      def clipWhenLowerLimitIsLessThanHigher(outputScaledValue, outputRange):
          if (outputScaledValue < outputRange[0]):
              return outputRange[0]
          elif (outputScaledValue > outputRange[1]):
              return outputRange[1]
          else:
              return outputScaledValue
          end
      end

      slope = computeSlope(rawRange, scaledRange)
      intercept = computeIntercept(slope, rawRange, scaledRange)
      scaledValue = slope * value + intercept
      return clipScaledValue(scaledValue, scaledRange)
  end

  def limit(value, range):
      return scale(value, range, range)
  end


  rq_init_comm_if_connected(9, "1")
  rq_init_comm_if_connected(2, "2")
  rq_init_comm_if_connected(3, "3")
  rq_init_comm_if_connected(4, "4")
  rq_print_connected_grippers()
  rq_gripper_communication_thread = run rq_gripper_communication()
  set_closed_norm(97.6470588235294, 1)
  set_open_norm(1.1764705882352942, 1)
  set_closed_mm(0.0, 1)
  set_open_mm(53.0, 1)
  set_closed_norm(100.0, 2)
  set_open_norm(0.0, 2)
  set_closed_mm(0.0, 2)
  set_open_mm(50.0, 2)
  set_closed_norm(100.0, 3)
  set_open_norm(0.0, 3)
  set_closed_mm(0.0, 3)
  set_open_mm(50.0, 3)
  set_closed_norm(100.0, 4)
  set_open_norm(0.0, 4)
  set_closed_mm(0.0, 4)
  set_open_mm(50.0, 4)
  rq_current_limit_enabled = False
  while(not rq_gripper_communication_thread_started):
      sync()
  end
  # end: URCap Installation Node
  # begin: URCap Installation Node
  #   Source: OPC UA, 2.0.2, Rocketfarm AS
  #   Type: OPC UA
  global opcua_daemon = rpc_factory("xmlrpc", "http://127.0.0.1:40409/RPC2")
  def opcua_client_connect(address):
  return opcua_daemon.client_connect(address)
  end
  def opcua_client_get_id(client_name):
  return opcua_daemon.client_get_id(client_name)
  end
  def opcua_client_try_connect(client_id):
  opcua_result = False
  if (opcua_daemon.client_connect(client_id)):
  sleep(0.01)
  opcua_result = opcua_daemon.client_is_connected(client_id)
  opcua_retry = 10
  while ( (not opcua_result) and (opcua_retry > 0) ):
  sleep(0.1)
  opcua_result = opcua_daemon.client_is_connected(client_id)
  opcua_retry = opcua_retry - 1
  end
  end
  return opcua_result
  end
  def opcua_client_disconnect(client_id):
  return opcua_daemon.client_disconnect(client_id)
  end
  def opcua_client_is_connected(client_id):
  return opcua_daemon.client_is_connected(client_id)
  end
  def opcua_client_read_byid(client_id, namespace_id, variable_id):
  return opcua_daemon.client_read_variable_by_id(client_id, namespace_id, variable_id)
  end
  def opcua_client_read_byname(client_id, namespace_id, variable_name):
  return opcua_daemon.client_read_variable_by_name(client_id, namespace_id, variable_name)
  end
  def opcua_client_write_byid(client_id, namespace_id, variable_id, variable_value):
  return opcua_daemon.client_write_variable_by_id(client_id, namespace_id, variable_id, variable_value)
  end
  def opcua_client_write_byname(client_id, namespace_id, variable_name, variable_value):
  return opcua_daemon.client_write_variable_by_name(client_id, namespace_id, variable_name, variable_value)
  end
  def opcua_client_last_error(client_id):
  return opcua_daemon.client_get_last_error(client_id)
  end
  def opcua_server_read_byname(variable_name):
  return opcua_daemon.server_read_variable_by_name(variable_name)
  end
  def opcua_server_write_byname(variable_name, variable_value):
  return opcua_daemon.server_write_variable_by_name(variable_name, variable_value)
  end
  def opcua_server_last_error():
  return opcua_daemon.server_get_last_error()
  end
  def opcua_error_to_string(errorCode):
  return opcua_daemon.error_code_to_string(errorCode)
  end
  # end: URCap Installation Node
  global AMR_Position=struct(position_identifier=0, x1=0, x2=0, y1=0, y2=0, theta1=0, theta2=0)
  global CAM_Pose=p[0,0,0,0,0,0]
  global CAM_Relation=""
  global CMD_Abort=  False
  global CMD_Clear=  False
  global CMD_Reset=  False
  global CMD_Start=  False
  global CMD_Suspend=  False
  global CMD_Unhold=  False
  global CMD_Unsuspend=  False
  global CNT_Rack_Output=0
  global FNC_Freedrive=  False
  global PRC_TubCounter=0
  global STP=0
  global easyPickCount=0
  global easyPickCount_4=0
  global easyPickCount_6=0
  global easyPickCount_7=0
  global easyPickNoObj=0
  global easyPickNoObj_4=0
  global easyPickNoObj_6=0
  global easyPickNoObj_7=0
  global easyPickParts=0
  global easyPickParts_4=0
  global easyPickParts_6=0
  global easyPickParts_7=0
  global Container_mid_1_p=p[-.379239199143, -.127191311915, .299999999998, .000000000046, -.000000000021, -1.247199999994]
  global Container_mid_1_q=[-2.477408934449926, -1.2969853503591224, -1.875639182904262, -1.539621866126728, 1.5731943360401213, -2.8009955944022717]
  global Container_capt_p=p[-.525590029047, .407247642794, .411588185841, -.000000000107, .000000000065, -2.896148821900]
  global Container_capt_q=[-3.5968351615224767, -2.0050156108707204, -0.8176271154495112, -1.8895759482008394, 1.5730967555598792, -2.2743681102957645]
  global Waypoint_51_p=p[-.335468094724, -.217855817953, .299999999998, .000000000047, -.000000000014, -.994837065669]
  global Waypoint_51_q=[-2.2250460001249586, -1.2969853503591224, -1.875639182904262, -1.539621866126728, 1.573194336040121, -2.800995594402271]
  global Waypoint_13_p=p[-.479450777041, .284140798427, .125270103493, -.276792173670, 2.098433187455, -2.121256516887]
  global Waypoint_13_q=[-2.8915050665484827, -1.9549266300597132, -2.2318272590637207, -1.6654960117735804, 0.020810842514038086, -0.4019392172442835]
  global Waypoint_70_p=p[-.472820924464, .292439826304, .207418370234, -.259787347864, -2.053484648504, 2.070709755662]
  global Waypoint_70_q=[-2.969927421603815, -2.07168115810532, -1.6835546062719366, -2.4953958198513964, 0.4489790927922641, -0.005578998612037367]
  global Waypoint_2_p=p[-.312961047461, -.152991312519, .223609826854, -.745314530454, -1.713873240489, 1.673341715282]
  global Waypoint_2_q=[-2.3560472170459192, -2.183784624139303, -1.4583134651184082, -2.6435262165465296, 1.6522362232208252, 0.043451953679323196]
  global Waypoint_3_p=p[-.113749865836, -.390110151572, .317307487562, -.519383711706, -.839884211339, 1.756868173041]
  global Waypoint_3_q=[-1.8909733931170862, -1.720626016656393, -1.5115610361099243, -2.1240560017027796, 2.1809096336364746, 0.7227501273155212]
  global Waypoint_15_p=p[.029144035010, -.436802470887, .327885032028, -.521560953301, -.623641814548, 1.862659450154]
  global Waypoint_15_q=[-1.564817253743307, -1.556895188321807, -1.6826975345611572, -1.6944714985289515, 2.2362685203552246, 1.117417335510254]
  global Waypoint_14_p=p[.068712235638, -.569419545175, .285215357659, -.679242949116, -.712065334485, 1.394044574094]
  global Waypoint_14_q=[-1.5731792953485346, -1.8029235103747094, -1.6781008808776736, -1.2218450646111982, 2.4719572998240125, 1.6394218026856375]
  global Waypoint_4_p=p[-.047220457210, -.557624911767, .136370962514, -.679242949107, -.712065334475, 1.394044574096]
  global Waypoint_4_q=[-1.7740079055958748, -2.0023561428872334, -1.7577251142892676, -1.18903287716154, 2.4487287370345143, 1.322902469273079]
  global Waypoint_25_p=p[.065436479647, -.569388431626, .287820755049, -.679242949185, -.712065334557, 1.394044574070]
  global Waypoint_25_q=[-1.5789263550890595, -1.8020194754825436, -1.6702557537748035, -1.237882536889547, 2.471995808083492, 1.6301087487321393]
  global Waypoint_39_p=p[.137772150180, -.577759956854, .299999999946, .000000000217, -.000000000207, -1.594351842625]
  global Waypoint_39_q=[-1.108978697428574, -1.776486680444405, -1.413737665315093, -1.5218908901738937, 1.5733062372356947, -1.0863866394180182]
  global Waypoint_41_p=p[.074222967010, -.565641640647, .234620140366, -.516884386806, .529223682286, -1.529619060506]
  global Waypoint_41_q=[-0.9596722604286052, -1.8767069964135548, -1.4892746174057256, -1.7813862040292285, 1.0520698599867686, -0.8199687448260349]
  global Waypoint_40_p=p[.039987741677, -.564832865048, .191055405868, -.767560686167, .343136533060, -2.241315728308]
  global Waypoint_40_q=[-1.0070649180116558, -1.8745927522477324, -1.6139175023195245, -1.6337474788493545, 1.032708081143138, -0.11587278312988403]
  global Waypoint_42_p=p[.041363380882, -.564865360786, .192805844739, .278500165520, .624117100927, .762272396553]
  global Waypoint_42_q=[-1.0050718976263102, -1.8744386685524779, -1.609151451954446, -1.6399653140247947, 1.0334006002355505, -3.254032861659603]
  global Waypoint_43_p=p[.041363380886, -.564865360780, .192805844755, .854271020883, .226833028600, 2.453002871494]
  global Waypoint_43_q=[-1.0050567614299233, -1.874341297657562, -1.6092945416026048, -1.6397580431809713, 1.0333661149462194, -5.0371728933995605]
  global Waypoint_44_p=p[.040882892233, -.564854254876, .192193763716, .110913882012, .659173708659, .275719738520]
  global Waypoint_44_q=[-1.0057704811530535, -1.8745207681598055, -1.6107765025572558, -1.637858394640876, 1.033164860873599, -2.7487836132940755]
  global Waypoint_45_p=p[.042647731639, -.564895808997, .194439423694, -.451694728506, .563172064821, -1.343350300184]
  global Waypoint_45_q=[-1.0032860829914387, -1.8741561795270565, -1.6048483308761785, -1.6453689714776623, 1.0342050634514657, -1.06078829880322]
  global Waypoint_46_p=p[.099944144487, -.566244126804, .267342790130, -.451694834765, .563172023386, -1.343350532536]
  global Waypoint_46_q=[-0.9257438092434924, -1.889970530402497, -1.3828165217629076, -1.8916791100652528, 1.0664350961373816, -0.9805910833329659]
  global Waypoint_47_p=p[.099944144444, -.566244126727, .267342790273, -.101742139519, .058679218003, -1.457888523314]
  global Waypoint_47_q=[-1.1112623176383014, -1.729989471869196, -1.5530029871033957, -1.4442770617454777, 1.4670579052775654, -1.2224020460061675]
  global Waypoint_48_p=p[-.136182767566, -.647487115908, .294247768372, -.101742139549, .058679218020, -1.457888523312]
  global Waypoint_48_q=[-1.532196177857717, -1.9115932455375173, -1.2651848069729779, -1.5055651746702665, 1.4703193777418382, -1.646379689188814]
  global Waypoint_49_p=p[-.159024328559, -.641021381179, .047691706070, -.000000000033, -.000000000027, -1.457897102937]
  global Waypoint_49_q=[-1.6098490079965062, -2.1164987141784586, -1.6156631902166785, -0.9800092198841526, 1.573231151532669, -1.722204302767242]
  global Waypoint_50_p=p[-.159024328558, -.641021381151, .291114489351, -.000000000033, -.000000000027, -1.457897102937]
  global Waypoint_50_q=[-1.609190265995684, -1.9426985888940234, -1.2189094859258596, -1.55056435122874, 1.5734384912955113, -1.7235116759964022]
  global Waypoint_53_p=p[-.050111345339, -.357608435610, .335880801283, .034180375734, .020280946727, -.284888945062]
  global Waypoint_53_q=[-1.3262308189700454, -1.2221767968893875, -1.8246061249803773, -1.7046285947349489, 1.567288986353525, -2.612420684434543]
  global Spatula_above_p=p[.241880327671, -.243077591927, .290283157642, .000026293989, -.000477463062, 3.067686800856]
  global Spatula_above_q=[-0.3881264518731289, -1.1433094134493045, -1.996913957798169, -1.572030383936684, 1.5734346414190374, 1.2567789862982233]
  global Spatula_pick_p=p[.240292635430, -.243077591534, .189212061148, .000026293987, -.000477463065, 3.067686800855]
  global Spatula_pick_q=[-0.39083408330539005, -1.1777602778656497, -2.2383115866577645, -1.2961817529600745, 1.573403050820434, 1.2551372216266965]
  global container_start_p=p[.200650292946, -.570238751958, .366326773614, 1.360500828661, .021700128770, 2.681649891414]
  global container_start_q=[-0.7669977765142582, -2.188996679669204, -0.7412727239230232, -2.581362891432544, 1.0193601740278728, 1.1884911920528847]
  global container_wp_1_p=p[.170613637794, -.572150573676, .294509026043, 1.259497117139, -.008270589399, 2.787717865625]
  global container_wp_1_q=[-0.8129253370121727, -2.0726598902108755, -1.0846040680899218, -2.2403146195823957, 1.0281191187839607, 1.0435744211830564]
  global Waypoint_55_p=p[.077280900603, -.567308602990, .212067617714, 1.259497117148, -.008270589399, 2.787717865619]
  global Waypoint_55_q=[-0.9181858327853867, -1.9744793804952083, -1.4540279077890048, -1.9155621911627945, 0.9643238328181578, 0.9457250675800015]
  global Waypoint_56_p=p[.135568164031, -.570867938153, .245215470413, 1.476861317558, -.018269607491, 2.679642659499]
  global Waypoint_56_q=[-0.8259784040282607, -2.108036981522602, -1.2111990877342924, -2.2405969375728745, 0.9451797152137279, 1.125710531287379]
  global Waypoint_74_p=p[.164827890887, -.574638012411, .193751361296, 2.053636896063, -.046507887560, 2.274278266449]
  global Waypoint_74_q=[-0.7657213433975762, -2.450387120010788, -0.9886183070290357, -2.7078095590939375, 0.8831550681477878, 1.5106229631053527]
  global ftr_scoop2_p=p[.194287054614, -.495779761333, .282072128495, -.179029871953, 1.612108092436, -.016025695011]
  global ftr_scoop2_q=[-0.5957383150173561, -2.264100500923713, -1.1936887184643812, -2.8893702964346097, 0.8750688478879766, -1.4109843517598684]
  global aftr_scoo3_p=p[-.289759911340, -.315385007342, .303743796282, .159961590809, 1.627415489603, -.344855744095]
  global aftr_scoo3_q=[-1.3374747909924949, -1.6809733407851706, -1.9857606509106667, -2.713564895186775, 0.5589807453366573, -1.3631067603374376]
  global Waypoint_60_p=p[-.013316432876, -.544772031582, .383371643081, 2.208233379808, .037543335712, 2.097559881761]
  global Waypoint_60_q=[-0.9328326161883087, -2.0999933666355775, -1.1958015693111372, -3.060905141293654, 0.690378518537611, 1.7121940951337198]
  global Waypoint_61_p=p[-.412188693372, -.356446875193, .383371643081, 1.751740964455, -.739956256289, 1.600691174920]
  global Waypoint_61_q=[-1.766185342973321, -2.0999933666355775, -1.1958015693111372, -3.060905141293654, 0.690378518537611, 1.7121940951337198]
  global Waypoint_75_p=p[-.343126484123, -.342779621892, .335357223804, .359429517288, 1.600352990741, -.365083732359]
  global Waypoint_75_q=[-1.517806275013295, -1.8136828056045395, -1.737638081810795, -2.8432599585466436, 0.5149430839716123, -1.4579122147201877]
  global aftr_scoop1_p=p[.138503854266, -.514479969882, .214153672011, -.134825326227, 1.559916297527, -.059196589314]
  global aftr_scoop1_q=[-0.6880464314785328, -2.2689986529709643, -1.3310176475983653, -2.673087158390708, 0.8340516295138949, -1.4557846480003231]
  global After_disp_3_p=p[.125934854156, -.585611107804, .299545938076, .959554236104, -.134386766509, 2.880651774211]
  global After_disp_3_q=[-0.9434480594885066, -2.016473586333989, -1.1036579072158617, -2.096459283015281, 1.1479556364931514, 0.8433331387406042]
  global Waypoint_62_p=p[-.542658707241, -.114281911009, .251261544113, 1.813043609523, -.679411528034, 1.655271622964]
  global Waypoint_62_q=[-2.158300033470912, -1.9418836862428677, -1.8142999147147894, -2.778920736683023, 0.21900622104017292, 1.8983390235012934]
  global Waypoint_63_p=p[.101294795191, -.465376052375, .381756220355, .972633305146, -.158447626639, 2.887199602585]
  global Waypoint_63_q=[-0.8528172446194038, -1.7393709485118478, -1.2544079521837954, -2.2703112963960628, 1.1965892397133469, 0.91867216443391]
  global Start_p=p[-.033064633790, -.365398531763, .389873206922, .000000000001, .000000000001, 2.725785203584]
  global Start_q=[-1.287596562866887, -1.232866726886848, -1.6880113260231102, -1.7912103151657988, 1.5729028131945846, 0.6981423183093938]
  global Waypoint_76_p=p[-.479450777041, .284140798427, .125270103493, -.276792173670, 2.098433187454, -2.121256516887]
  global Waypoint_76_q=[-2.891505066548503, -1.9549266300590151, -2.231827259067863, -1.6654960117542226, 0.020810842514162875, -0.4019392172601952]
  global PowderA_wayp1_p=p[-.472820924474, .292439826233, .207418370237, -.137787250486, 2.177332259632, -2.152029714756]
  global PowderA_wayp1_q=[-2.911134078210732, -1.90240864358569, -1.968768330510411, -2.500365101593811, 0.11427687110891149, 0.0958980389250167]
  global Waypoint_80_p=p[-.303921889165, -.326082520111, .297721580072, -.584846481381, 1.914382606328, -1.960922301253]
  global Waypoint_80_q=[-1.6364180099980672, -2.041258366871811, -1.472153549517767, -2.7572808013122696, 0.9684003593854582, 0.047163023020230455]
  global Decapp_above_p=p[-.013480295948, -.359153355979, .266194408367, -.879653555922, 1.646336924805, -1.709111068605]
  global Decapp_above_q=[-0.9632157249872035, -2.0163405763031657, -1.5968194594157152, -2.6579215719847085, 1.251243398585566, 0.047906446502667066]
  global Decapp_place_p=p[-.013480295848, -.359153356116, .158558645017, -.879653554904, 1.646336919751, -1.709111066446]
  global Decapp_place_q=[-0.9633419174801583, -2.157735564881908, -1.695182597572722, -2.418253553201909, 1.2517436353048952, 0.04819090596102882]
  global Waypoint_78_p=p[-.051450028091, -.519555688329, .365718563414, -1.287302938145, 1.077637394477, -1.218524965834]
  global Waypoint_78_q=[-0.9214276262416012, -1.8899696965062578, -1.4939326452510562, -2.840015661555725, 0.5585157189668353, 0.033997638875617575]
  global Waypoint_81_p=p[-.030847790230, -.346237542439, .241203613248, .000000000000, .000000000000, .000000000000]
  global Waypoint_81_q=[-1.265848516232941, -1.1652881302267932, -2.11003646605462, -1.4369228603041853, 1.573284436504383, -2.835929896730388]
  global Waypoint_79_p=p[-.030847972829, -.346235312674, .229874122470, .000000000000, .000000000000, .000000000000]
  global Waypoint_79_q=[-1.2659333103898618, -1.1699230683425625, -2.1365870669440055, -1.4057372655396474, 1.5732787836040316, -2.8358953794066757]
  global Waypoint_82_p=p[-.031079593487, -.346547394534, .293012696855, -.000011575267, -.000017731224, -.000713984074]
  global Waypoint_82_q=[-1.2664169521879751, -1.1572597700415788, -1.982185304253158, -1.5727862504184884, 1.5732673022058234, -2.83632822711502]
  global Cap_above_p=p[-.163602500478, -.618357694237, .258271116068, .000026793591, -.000032305852, -.969382601663]
  global Cap_above_q=[-1.6181634639269902, -1.896432778341337, -1.3662765317923142, -1.449515114018281, 1.5734416863575176, -2.220489512402157]
  global Cap_Place_p=p[-.153420247224, -.637174247221, .035295616791, .000000000002, -.000000000002, -1.457849918374]
  global Cap_Place_q=[-1.6014084627078784, -2.123124488207292, -1.6429187572395012, -0.946127085055064, 1.573175527437006, -1.7136981844648291]
  global OP_PowderA2_p=p[.009371277507, -.409434369247, .294169017766, -.823281033205, 1.709410851243, -1.698303593897]
  global OP_PowderA2_q=[-0.9994544761745754, -2.1395254572673217, -1.3437567783153916, -2.8143375616690456, 1.2617899549595724, 0.019614613715634555]
  global OP_PowderA_abov_p=p[-.012145216791, -.363335041455, .315325728178, -.777135478411, 1.752984823781, -1.740925591659]
  global OP_PowderA_abov_q=[-1.01634425044037, -2.024785947780374, -1.4658894155189923, -2.8070189735738786, 1.3091674480404514, 0.020022086766872782]
  global OP_PowderA_pick_p=p[-.012145216707, -.363335041590, .179898787547, -.777135478413, 1.752984823781, -1.740925591659]
  global OP_PowderA_pick_q=[-1.0165129229305911, -2.176980100858497, -1.6127054339661555, -2.5080740815244567, 1.3098787614888208, 0.020270375244195882]
  global Op_PowA_wP_p=p[-.173727579245, -.372934016396, .295116627479, -.972390492433, 1.540962074418, -1.548745344994]
  global Op_PowA_wP_q=[-1.1740587397768483, -1.865656321049359, -1.7426943793777419, -2.679427276872525, 0.8588908769087338, 0.017944699631825187]
  global Waypoint_1_p=p[-.451048883256, -.340589460864, .308223661552, .097058877504, .091048998701, -1.578386010942]
  global Waypoint_1_q=[-2.222400490437643, -1.7554131946959437, -1.398173213005066, -1.6564461193480433, 1.5042352676391602, -2.2106884161578577]
  global Spatula_otw_p=p[-.038472058237, -.263141484147, .425351216717, -.000441582511, -.000128175490, 3.034387645854]
  global Spatula_otw_q=[-1.1888947506684495, -1.0083288774886814, -1.7052227056065874, -1.9984805067363443, 1.5730180972985317, 0.48793409320312264]
  global pick_spat_L_abv_p=p[.247376339171, -.151300871293, .298405979617, .000026293989, -.000477463062, 3.067686800856]
  global pick_spat_L_abv_q=[-0.07082187843937948, -0.9918336120099029, -2.048431407771396, -1.6719226065707566, 1.5735148227092874, 1.5739821706892307]
  global spat_L_pick_p=p[.244425006707, -.151048053384, .192288246285, .000026293989, -.000477463065, 3.067686800855]
  global spat_L_pick_q=[-0.07170850917614935, -0.9939169317558161, -2.3190151588645502, -1.3992549297298966, 1.573619586467819, 1.5742112847515592]
  global spat_L_lift_p=p[.247500241215, -.151291104039, .242146826477, .000026293989, -.000477463064, 3.067686800855]
  global spat_L_lift_q=[-0.07132168213116863, -0.9873531406871798, -2.1938095635783172, -1.531024644535787, 1.5736129628476565, 1.5740661231239859]
  global spat_L_side_p=p[.251772314117, -.093610100391, .242165935204, .000026293989, -.000477463064, 3.067686800855]
  global spat_L_side_q=[0.16311920731341095, -0.9159674867544636, -2.2202625845173465, -1.5759061264106862, 1.5736725172206427, 1.8084579794657634]
  global spat_L_up_p=p[.248631729748, -.094370561652, .425351216716, .000026293989, -.000477463065, 3.067686800855]
  global spat_L_up_q=[0.16435650344985986, -1.008385469590376, -1.7051729211515223, -1.9985780211252369, 1.5729805495343943, 1.8078858605162342]
  global spat_M_up_p=p[.246651483123, -.200758466677, .427983242435, .000026293988, -.000477463066, 3.067686800854]
  global spat_M_up_q=[-0.2488061154947081, -1.1388154682286178, -1.6405006043284098, -1.932909670500866, 1.5729930693357987, 1.394694958078517]
  global spat_M_pick_p=p[.243754824031, -.195909855689, .192274495860, .000026293989, -.000477463063, 3.067686800855]
  global spat_M_pick_q=[-0.2371047546337337, -1.0815273547611497, -2.2806002623741977, -1.3500947192370933, 1.573515135501001, 1.4088438823663394]
  global spat_S_up_p=p[.250500617207, -.246905508589, .391583682111, .000026293987, -.000477463068, 3.067686800854]
  global spat_S_up_q=[-0.3880360419879594, -1.1962881911765244, -1.7058643812256875, -1.8101014540154097, 1.5731545967396166, 1.2558061200976702]
  global spat_S_pick_p=p[.245173607467, -.244249950907, .193022226997, .000026293988, -.000477463064, 3.067686800854]
  global spat_S_pick_q=[-0.38836215799357987, -1.1880037605751017, -2.222350098157584, -1.30189927792612, 1.5733998957551099, 1.2575641527417636]
  def Sub_Vision_V18():
    $ 732 "Sub_Vision_V18" "noBreak"
    $ 733 "PreSettings"
    $ 734 "CAM_LM_Detected≔ False "
    global CAM_LM_Detected=  False
    $ 735 "CAM_Captures≔0"
    global CAM_Captures=0
    $ 736 "CAM_Pose≔p[0,0,0,0,0,0]"
    global CAM_Pose=p[0,0,0,0,0,0]
    $ 737 "CAM_LM_Refinmnt≔ False "
    global CAM_LM_Refinmnt=  False
    $ 738 "CAM_LM_Refined≔ False "
    global CAM_LM_Refined=  False
    $ 739 "CAM_LM_Deviatn≔p[0,0,0,0,0,0]"
    global CAM_LM_Deviatn=p[0,0,0,0,0,0]
    $ 740 "CAM_LM_ID≔0"
    global CAM_LM_ID=0
    $ 741 "CAM_Done≔ False "
    global CAM_Done=  False
    $ 742 "CAM_CNT_Obj≔0"
    global CAM_CNT_Obj=0
    $ 743 "CAM_Result = []"
    CAM_Result = []
    $ 744 "OBJ_Detected≔ False "
    global OBJ_Detected=  False
    $ 745 "FRM_Reference≔p[0,0,0,0,0,0]"
    global FRM_Reference=p[0,0,0,0,0,0]
    $ 746 "'=========='"
    # '=========='
    $ 747 "Switch Action"
    switch_1 = Action
    $ 748 "Case 13"
    if (13 == switch_1):
    elif (15 == switch_1):
      $ 866 "Case 15"
    elif (131 == switch_1):
      $ 912 "Case 131"
      $ 913 "Read (SensoPart)"
      $ 914 "Action_Info≔'search for landmark'"
      global Action_Info="search for landmark"
      $ 915 "CAM_LM≔CAM_LMs[4]"
      global CAM_LM=CAM_LMs[4]
      $ 916 "CAM_Relation≔CAM_LM.capture_relation"
      global CAM_Relation=CAM_LM.capture_relation
      $ 917 "go to capture pose"
      $ 920 "If ITM_ID≟1 and JIG≟7"
      if (ITM_ID == 1  and  JIG == 7):
        $ 921 "PSE_T≔uLM_Cap_SSRack"
        global PSE_T=uLM_Cap_SSRack
      else:
        $ 922 "ElseIf ITM_ID≟5 and JIG≟7"
        if (ITM_ID == 5  and  JIG == 7):
          $ 923 "PSE_T≔FRM_Cap_SSRack"
          global PSE_T=FRM_Cap_SSRack
        else:
          $ 924 "ElseIf ITM_ID≟13 and JIG≟7"
          if (ITM_ID == 13  and  JIG == 7):
            $ 925 "PSE_T≔FRM_pick_rack_const"
            global PSE_T=p[-0.5568395192387274,0.34423986364170267,0.44698620470146266,-1.0069110132199915E-6,3.378712467497258E-5,-8.002029546773325E-6]
          else:
            $ 926 "ElseIf ITM_ID≟1 and JIG≟15"
            if (ITM_ID == 1 and JIG == 15):
              $ 927 "MoveJ"
              $ 928 "Container_mid_1" "breakAfter"
              movej(get_inverse_kin(Container_mid_1_p, qnear=Container_mid_1_q), a=1.3962634015954636, v=1.0471975511965976, r=0.05)
              $ 929 "Container_capt" "breakAfter"
              movej(get_inverse_kin(Container_capt_p, qnear=Container_capt_q), a=1.3962634015954636, v=1.0471975511965976)
              $ 930 "PSE_T≔FRM_Container_S_const"
              global PSE_T=p[-0.510412665574981,0.40064363362973565,0.41159789496794374,-1.1370875604168537E-5,-3.643547521609506E-6,-2.896122366208473]
            else:
              $ 931 "ElseIf ITM_ID≟1 and JIG≟16"
              if (ITM_ID == 1  and  JIG == 16):
                $ 932 "MoveJ"
                $ 933 "Waypoint_51" "breakAfter"
                movej(get_inverse_kin(Waypoint_51_p, qnear=Waypoint_51_q), a=1.3962634015954636, v=1.0471975511965976, r=0.05)
                $ 935 "PSE_T≔FRM_Weigh_scale_const"
                global PSE_T=p[-0.3454891122972868,0.06305469656946562,0.547028193804949,1.63274868305228E-4,-7.686242288056818E-5,-2.2741025165393225]
              else:
                $ 936 "ElseIf ITM_ID≟1 and JIG≟17"
                if (ITM_ID == 1  and  JIG == 17):
                  $ 937 "MoveJ"
                  $ 938 "Waypoint_51" "breakAfter"
                  movej(get_inverse_kin(Waypoint_51_p, qnear=Waypoint_51_q), a=1.3962634015954636, v=1.0471975511965976, r=0.05)
                  $ 940 "PSE_T≔FRM_Weigh_scale_const"
                  global PSE_T=p[-0.3454891122972868,0.06305469656946562,0.547028193804949,1.63274868305228E-4,-7.686242288056818E-5,-2.2741025165393225]
                else:
                  $ 941 "ElseIf ITM_ID≟1 and JIG≟21"
                  if (ITM_ID == 1  and  JIG == 21):
                    $ 942 "MoveJ"
                    $ 943 "Waypoint_51" "breakAfter"
                    movej(get_inverse_kin(Waypoint_51_p, qnear=Waypoint_51_q), a=1.3962634015954636, v=1.0471975511965976, r=0.05)
                    $ 945 "PSE_T≔FRM_PoTS_const"
                    global PSE_T=p[-0.5211683440725288,-0.17068665293155189,0.5469908617304544,2.009713344566374E-4,5.545167142016751E-6,-2.2342044673695503]
                  end
                end
              end
            end
          end
        end
      end
      $ 946 "do_transition(PSE_T, keep_rxry=False)"
      do_transition(PSE_T, keep_rxry=False)
      $ 947 "Set"
      set_tcp(p[0.0,0.0,0.161,3.1415,0.0,0.0])
      $ 948 "MoveJ"
      $ 949 "PSE_T" "breakAfter"
      movej(PSE_T, a=1.3962634015954636, v=1.7453292519943295)
      $ 950 "CAM_Pose≔get_actual_tcp_pose()"
      global CAM_Pose= get_actual_tcp_pose ()
      $ 951 "Loop  not CAM_Done and  not ERROR.FLAG and  not CMD_Stop"
      while (  not  CAM_Done  and    not  ERROR.FLAG  and    not  CMD_Stop):
        $ 952 "adjust capture pose"
        $ 953 "If CAM_LM_Detected and CAM_LM_Refinmnt"
        if (CAM_LM_Detected  and  CAM_LM_Refinmnt):
          $ 954 "PSE_T≔p[0,0,0.300,0,0,0]"
          global PSE_T=p[0,0,0.300,0,0,0]
          $ 955 "CAM_Pose≔PSE_T"
          global CAM_Pose=PSE_T
          $ 956 "If  not is_reachable(FRM_Reference,[PSE_T])"
          if (  not  is_reachable(FRM_Reference,[PSE_T])):
            $ 957 "Error"
            $ 958 "set_error(ERROR_POSE_NOT_REACHABLE)"
            set_error(ERROR_POSE_NOT_REACHABLE)
          end
          $ 959 "If  not ERROR.FLAG"
          if (  not  ERROR.FLAG):
            $ 960 "MoveJ"
            $ 961 "PSE_T" "breakAfter"
            set_tcp(p[0.0,0.0,0.161,0.0,0.0,0.0])
            movej(pose_trans(FRM_Reference, PSE_T), a=0.8726646259971648, v=1.3962634015954636)
            $ 962 "CAM_LM_Refined≔ True "
            global CAM_LM_Refined=  True
          end
        else:
          $ 963 "ElseIf  not CAM_LM_Detected and CAM_Captures>0"
          if (  not  CAM_LM_Detected  and  CAM_Captures>0):
            $ 964 "MoveL"
            $ 965 "If FRM_Reference≟p[0,0,0,0,0,0]"
            if (FRM_Reference == p[0,0,0,0,0,0]):
              $ 966 "PSE_T≔get_random_pose(pose_ref=CAM_Pose, mode='cubic', range_max=[0.150,0.150,0.015])"
              global PSE_T=get_random_pose(pose_ref=CAM_Pose, mode="cubic", range_max=[0.150,0.150,0.015])
            else:
              $ 971 "Else" "noBreak"
              $ 972 "PSE_T≔get_random_pose(pose_ref=CAM_Pose, mode='rotation', range_max=[10,10,0])"
              global PSE_T=get_random_pose(pose_ref=CAM_Pose, mode="rotation", range_max=[10,10,0])
              $ 973 "CAM_LM_Refined≔ True "
              global CAM_LM_Refined=  True
            end
            $ 974 "If get_inverse_kin_has_solution(pose_trans(FRM_Reference, PSE_T))"
            if (get_inverse_kin_has_solution( pose_trans (FRM_Reference, PSE_T))):
              $ 975 "Comment"
              # Comment
              $ 976 "PSE_T" "breakAfter"
              set_tcp(p[0.0,0.0,0.161,3.1415,0.0,0.0])
              movel(pose_trans(FRM_Reference, PSE_T), a=0.03, v=0.05)
            else:
              $ 977 "Else" "noBreak"
              $ 978 "'If random pose is out of reach, set the initial cam pose'"
              # 'If random pose is out of reach, set the initial cam pose'
              $ 979 "PSE_T≔CAM_Pose"
              global PSE_T=CAM_Pose
            end
          end
        end
        $ 980 "Wait: 2.0"
        sleep(2.0)
        $ 981 "trigger"
        $ 982 "If ITM_ID≟1 and JIG≟7"
        if (ITM_ID == 1  and  JIG == 7):
          # begin: URCap Program Node
          #   Source: SensoPart VISOR Robotic, 2.0.0, SensoPart Industriesensorik GmbH
          #   Type: VISOR Trigger
          $ 983 "# 1 VISOR Trigger"
          visor_changeJob(1, "Landmark_INVITE_2", 6000)
          visor_trigger(1, 6000, "arm")
          # end: URCap Program Node
        else:
          $ 984 "ElseIf ITM_ID≟5 and JIG≟7"
          if (ITM_ID == 5  and  JIG == 7):
            # begin: URCap Program Node
            #   Source: SensoPart VISOR Robotic, 2.0.0, SensoPart Industriesensorik GmbH
            #   Type: VISOR Trigger
            $ 985 "# 1 VISOR Trigger"
            visor_changeJob(1, "Landmark_INVITE_2", 6000)
            visor_trigger(1, 6000, "arm")
            # end: URCap Program Node
          else:
            $ 986 "ElseIf ITM_ID≟13 and JIG≟7"
            if (ITM_ID == 13  and  JIG == 7):
              # begin: URCap Program Node
              #   Source: SensoPart VISOR Robotic, 2.0.0, SensoPart Industriesensorik GmbH
              #   Type: VISOR Trigger
              $ 987 "# 1 VISOR Trigger"
              visor_changeJob(1, "Landmark_INVITE_2", 6000)
              visor_trigger(1, 6000, "arm")
              # end: URCap Program Node
            else:
              $ 988 "ElseIf ITM_ID≟1 and JIG≟15"
              if (ITM_ID == 1 and JIG == 15):
                # begin: URCap Program Node
                #   Source: SensoPart VISOR Robotic, 2.0.0, SensoPart Industriesensorik GmbH
                #   Type: VISOR Trigger
                $ 989 "# 1 VISOR Trigger"
                visor_changeJob(1, "PowderA", 6000)
                visor_trigger(1, 6000, "arm")
                # end: URCap Program Node
              else:
                $ 990 "ElseIf ITM_ID≟1 and JIG≟16"
                if (ITM_ID == 1 and JIG == 16):
                  # begin: URCap Program Node
                  #   Source: SensoPart VISOR Robotic, 2.0.0, SensoPart Industriesensorik GmbH
                  #   Type: VISOR Trigger
                  $ 991 "# 1 VISOR Trigger"
                  visor_changeJob(1, "Weigh_target", 6000)
                  visor_trigger(1, 6000, "arm")
                  # end: URCap Program Node
                else:
                  $ 992 "ElseIf ITM_ID≟1 and JIG≟17"
                  if (ITM_ID == 1 and JIG == 17):
                    # begin: URCap Program Node
                    #   Source: SensoPart VISOR Robotic, 2.0.0, SensoPart Industriesensorik GmbH
                    #   Type: VISOR Trigger
                    $ 993 "# 1 VISOR Trigger"
                    visor_changeJob(1, "Weigh_target", 6000)
                    visor_trigger(1, 6000, "arm")
                    # end: URCap Program Node
                  else:
                    $ 994 "ElseIf ITM_ID≟1 and JIG≟21"
                    if (ITM_ID == 1 and JIG == 21):
                      # begin: URCap Program Node
                      #   Source: SensoPart VISOR Robotic, 2.0.0, SensoPart Industriesensorik GmbH
                      #   Type: VISOR Trigger
                      $ 995 "# 1 VISOR Trigger"
                      visor_changeJob(1, "Weigh_target", 6000)
                      visor_trigger(1, 6000, "arm")
                      # end: URCap Program Node
                    end
                  end
                end
              end
            end
          end
        end
        $ 999 "TM_3D_Found≔visor_partsFound(1)"
        global TM_3D_Found= visor_partsFound (1)
        $ 1000 "If TM_3D_Found>0"
        if (TM_3D_Found>0):
          $ 1001 "CAM_LM_Detected≔ True "
          global CAM_LM_Detected=  True
          $ 1002 "CAM_Captures≔0"
          global CAM_Captures=0
        else:
          $ 1003 "Else" "noBreak"
          $ 1004 "CAM_LM_Detected≔ False "
          global CAM_LM_Detected=  False
          $ 1005 "CAM_Captures≔CAM_Captures+1"
          global CAM_Captures=CAM_Captures+1
        end
        $ 1010 "result"
        $ 1011 "If CAM_LM_Detected"
        if (CAM_LM_Detected):
          $ 1012 "If (CAM_LM_Refinmnt and CAM_LM_Refined) or  not CAM_LM_Refinmnt"
          if ((CAM_LM_Refinmnt  and  CAM_LM_Refined)  or    not  CAM_LM_Refinmnt):
            $ 1070 "If ITM_ID≟1 and JIG≟7"
            if (ITM_ID == 1  and  JIG == 7):
              $ 1071 "CAM_LM_SSRack≔visor_getPose3d(1, 0)"
              global CAM_LM_SSRack= visor_getPose3d (1, 0)
            else:
              $ 1072 "ElseIf ITM_ID≟5 and JIG≟7"
              if (ITM_ID == 5  and  JIG == 7):
                $ 1073 "CAM_LM_SSRack≔visor_getPose3d(1, 0)"
                global CAM_LM_SSRack= visor_getPose3d (1, 0)
              else:
                $ 1074 "ElseIf ITM_ID≟13 and JIG≟7"
                if (ITM_ID == 13  and  JIG == 7):
                  $ 1075 "CAM_LM_Bott≔visor_getPose3d(1, 0)"
                  global CAM_LM_Bott= visor_getPose3d (1, 0)
                else:
                  $ 1076 "ElseIf ITM_ID≟1 and JIG≟15"
                  if (ITM_ID == 1 and JIG == 15):
                    $ 1077 "CAM_LM_Cont_S≔visor_getPose3d(1, 0)"
                    global CAM_LM_Cont_S= visor_getPose3d (1, 0)
                    $ 1078 "cont_img_pose≔get_actual_tcp_pose()"
                    global cont_img_pose= get_actual_tcp_pose ()
                  else:
                    $ 1079 "ElseIf ITM_ID≟1 and JIG≟16"
                    if (ITM_ID == 1 and JIG == 16):
                      $ 1080 "CAM_cont≔visor_getPose3d(1, 0)"
                      global CAM_cont= visor_getPose3d (1, 0)
                      $ 1081 "cont_img_pose≔get_actual_tcp_pose()"
                      global cont_img_pose= get_actual_tcp_pose ()
                    else:
                      $ 1082 "ElseIf ITM_ID≟1 and JIG≟17"
                      if (ITM_ID == 1 and JIG == 17):
                        $ 1084 "cont_img_pose≔get_actual_tcp_pose()"
                        global cont_img_pose= get_actual_tcp_pose ()
                      else:
                        $ 1085 "ElseIf ITM_ID≟1 and JIG≟21"
                        if (ITM_ID == 1 and JIG == 21):
                          $ 1087 "cont_img_pose≔get_actual_tcp_pose()"
                          global cont_img_pose= get_actual_tcp_pose ()
                        end
                      end
                    end
                  end
                end
              end
            end
            $ 1088 "CAM_Done≔ True "
            global CAM_Done=  True
          end
        else:
          $ 1089 "ElseIf  not CAM_LM_Detected and CAM_Captures<CAM_PRM_Retries"
          if (  not  CAM_LM_Detected  and  CAM_Captures<CAM_PRM_Retries):
            $ 1090 "CAM_LM_Refined≔ False "
            global CAM_LM_Refined=  False
          else:
            $ 1091 "ElseIf CAM_Captures≥CAM_PRM_Retries"
            if (CAM_Captures >= CAM_PRM_Retries):
              $ 1092 "CAM_Done≔ True "
              global CAM_Done=  True
              $ 1093 "Error"
              $ 1094 "set_error(ERROR_NO_LANDMARK)"
              set_error(ERROR_NO_LANDMARK)
            end
          end
        end
      end
    elif (151 == switch_1):
      $ 1095 "Case 151"
      $ 1096 "Detect (SensoPart)"
      $ 1097 "go to capture pose"
      $ 1098 "FRM_Reference≔FRM_Cap_SSRack"
      global FRM_Reference=FRM_Cap_SSRack
      $ 1099 "PSE_T≔p[0,0,-0.00,0,0,0]"
      global PSE_T=p[0,0,-0.00,0,0,0]
      $ 1100 "do_transition(pose_trans(FRM_Reference, PSE_T), keep_rxry=False)"
      do_transition( pose_trans (FRM_Reference, PSE_T), keep_rxry=False)
      $ 1101 "JNT_Q≔get_actual_joint_positions()"
      global JNT_Q= get_actual_joint_positions ()
      $ 1102 "JNT_Q≔[JNT_Q[0], JNT_Q[1], JNT_Q[2], JNT_Q[3], JNT_Q[4], 0]"
      global JNT_Q=[JNT_Q[0], JNT_Q[1], JNT_Q[2], JNT_Q[3], JNT_Q[4], 0]
      $ 1103 "Set"
      set_tcp(p[0.0,0.0,0.161,3.1415,0.0,0.0])
      $ 1104 "movej(get_inverse_kin(pose_trans(FRM_Reference, PSE_T), qnear=JNT_Q))"
      movej(get_inverse_kin( pose_trans (FRM_Reference, PSE_T), qnear=JNT_Q))
      $ 1105 "CAM_Pose≔pose_trans(pose_inv(FRM_Reference), get_actual_tcp_pose())"
      global CAM_Pose= pose_trans ( pose_inv (FRM_Reference),  get_actual_tcp_pose ())
      $ 1106 "Loop  not CAM_Done and  not ERROR.FLAG and  not CMD_Stop"
      while (  not  CAM_Done  and    not  ERROR.FLAG  and    not  CMD_Stop):
        $ 1107 "If  not OBJ_Detected and CAM_Captures>0"
        if (  not  OBJ_Detected  and  CAM_Captures>0):
          $ 1108 "MoveL"
          $ 1109 "If FRM_Reference≟p[0,0,0,0,0,0]"
          if (FRM_Reference == p[0,0,0,0,0,0]):
            $ 1111 "PSE_T≔get_random_pose(pose_ref=CAM_Pose, mode='rotation', range_max=[15,15,0])"
            global PSE_T=get_random_pose(pose_ref=CAM_Pose, mode="rotation", range_max=[15,15,0])
          else:
            $ 1112 "Else" "noBreak"
            $ 1113 "PSE_T≔get_random_pose(pose_ref=CAM_Pose, mode='rotation', range_max=[10,10,0])"
            global PSE_T=get_random_pose(pose_ref=CAM_Pose, mode="rotation", range_max=[10,10,0])
          end
          $ 1114 "If get_inverse_kin_has_solution(pose_trans(FRM_Reference, PSE_T))"
          if (get_inverse_kin_has_solution( pose_trans (FRM_Reference, PSE_T))):
            $ 1115 "PSE_T" "breakAfter"
            set_tcp(p[0.0,0.0,0.161,3.1415,0.0,0.0])
            movel(pose_trans(FRM_Reference, PSE_T), a=0.03, v=0.05)
          else:
            $ 1116 "Else" "noBreak"
            $ 1117 "'If random pose is out of reach, set the initial cam pose'"
            # 'If random pose is out of reach, set the initial cam pose'
            $ 1118 "PSE_T≔CAM_Pose"
            global PSE_T=CAM_Pose
            $ 1119 "PSE_T" "breakAfter"
            set_tcp(p[0.0,0.0,0.161,3.1415,0.0,0.0])
            movel(pose_trans(FRM_Reference, PSE_T), a=0.03, v=0.05)
          end
        end
        $ 1120 "Wait: 0.5"
        sleep(0.5)
        $ 1121 "Set"
        set_tcp(p[0.0,0.0,0.161,3.1415,0.0,0.0])
        # begin: URCap Program Node
        #   Source: SensoPart VISOR Robotic, 2.0.0, SensoPart Industriesensorik GmbH
        #   Type: VISOR Trigger
        $ 1122 "# 1 VISOR Trigger"
        visor_changeJob(1, "Object Detection Single", 6000)
        visor_trigger(1, 6000, "arm")
        # end: URCap Program Node
        $ 1123 "If visor_isResponseOk(1)"
        if ( visor_isResponseOk (1)):
          $ 1124 "CAM_CNT_Obj≔visor_partsFound(1)"
          global CAM_CNT_Obj= visor_partsFound (1)
          $ 1125 "CAM_OBJ_Pose≔visor_getPose3d(1, 0)"
          global CAM_OBJ_Pose= visor_getPose3d (1, 0)
          $ 1126 "If CAM_CNT_Obj>0"
          if (CAM_CNT_Obj>0):
            $ 1127 "CAM_OBJ_Color≔visor_getAdditionalData(1, 0)"
            global CAM_OBJ_Color= visor_getAdditionalData (1, 0)
            $ 1128 "CAM_DetectScore≔to_num(visor_getAdditionalData(1, 1))/1000"
            global CAM_DetectScore=to_num( visor_getAdditionalData (1, 1))/1000
            $ 1129 "OBJ_Detected≔ True "
            global OBJ_Detected=  True
          end
        else:
          $ 1130 "Else" "noBreak"
          $ 1131 "CAM_Captures≔CAM_Captures+1"
          global CAM_Captures=CAM_Captures+1
        end
        $ 1132 "If OBJ_Detected"
        if (OBJ_Detected):
          $ 1133 "Get object data"
          $ 1134 "PRC_CntDetect≔0"
          global PRC_CntDetect=0
          $ 1135 "Loop PRC_CntDetect<CAM_CNT_Obj"
          while (PRC_CntDetect<CAM_CNT_Obj):
            $ 1136 "get object and jig number"
            $ 1137 "If ITM_ID≟1 and JIG≟7"
            if (ITM_ID == 1  and  JIG == 7):
              $ 1138 "FRM_Reference≔FRM_Cap_SSRack"
              global FRM_Reference=FRM_Cap_SSRack
            else:
              $ 1139 "ElseIf ITM_ID≟5 and JIG≟7"
              if (ITM_ID == 5  and  JIG == 7):
                $ 1140 "FRM_Reference≔uLM_Cap_SSRack"
                global FRM_Reference=uLM_Cap_SSRack
              end
            end
            $ 1143 "PSE_T≔pose_trans(pose_inv(FRM_Reference), CAM_OBJ_Pose)"
            global PSE_T= pose_trans ( pose_inv (FRM_Reference), CAM_OBJ_Pose)
            $ 1144 "CAM_Result.append(get_pattern_counter(PSE_T, 'X', pattern=[10, 5], patternsize=[0.181, 0.081]))"
            CAM_Result.append(get_pattern_counter(PSE_T, "X", pattern=[10, 5], patternsize=[0.181, 0.081]))
            $ 1145 "PRC_CntDetect≔PRC_CntDetect+1"
            global PRC_CntDetect=PRC_CntDetect+1
          end
          $ 1146 "CAM_Done≔ True "
          global CAM_Done=  True
        else:
          $ 1147 "ElseIf CAM_Captures≥CAM_PRM_Retries"
          if (CAM_Captures >= CAM_PRM_Retries):
            $ 1148 "CAM_Done≔ True "
            global CAM_Done=  True
          else:
            $ 1149 "Else" "noBreak"
            $ 1150 "CAM_Captures≔CAM_Captures+1"
            global CAM_Captures=CAM_Captures+1
          end
        end
      end
    end
    $ 1151 "'=========='"
    # '=========='
    $ 1152 "PostSettings"
    $ 1153 "FRM_Reference≔p[0,0,0,0,0,0]"
    global FRM_Reference=p[0,0,0,0,0,0]
    $ 1154 "Set"
    set_tcp(p[0.0,0.0,0.161,3.1415,0.0,0.0])
    $ 1155 "CAM_Pose≔p[0,0,0,0,0,0]"
    global CAM_Pose=p[0,0,0,0,0,0]
    $ 1156 "Action≔0"
    global Action=0
    $ 1157 "Action_Info≔''"
    global Action_Info=""
  end
  def Sub_AMR_MiR_V3():
    $ 1158 "Sub_AMR_MiR_V3" "noBreak"
    $ 1159 "PreSettings"
    $ 1160 "AMR_TargetList≔[1,2,3,4,5,21,22,23,24,31,32,33,34,35,36,37,38,41]"
    global AMR_TargetList=[1,2,3,4,5,21,22,23,24,31,32,33,34,35,36,37,38,41]
    $ 1161 "AMR_Done≔ False "
    global AMR_Done=  False
    $ 1162 "AMR_PosActual≔T2O_Current_Pos"
    global AMR_PosActual=modbus_get_signal_status("T2O_Current_Pos")
    $ 1163 "AMR_Attemps≔T2O_Nav_Attemps"
    global AMR_Attemps=modbus_get_signal_status("T2O_Nav_Attemps")
    $ 1164 "AMR_Battery≔MiR_Battery_Lvl"
    global AMR_Battery=modbus_get_signal_status("MiR_Battery_Lvl")
    $ 1165 "AMR_Charging≔(T2O_Charging≟1)"
    global AMR_Charging=(modbus_get_signal_status("T2O_Charging") == 1)
    $ 1166 "AMR_Position≔struct(position_identifier=T2O_Current_Pos, x1=MiR_Position_X1, x2=MiR_Position_X2, y1=MiR_Position_Y1, y2=MiR_Position_Y2, theta1=MiR_Theta_1, theta2=MiR_Theta_2) "
    global AMR_Position=struct(position_identifier=modbus_get_signal_status("T2O_Current_Pos"), x1=modbus_get_signal_status("MiR_Position_X1"), x2=modbus_get_signal_status("MiR_Position_X2"), y1=modbus_get_signal_status("MiR_Position_Y1"), y2=modbus_get_signal_status("MiR_Position_Y2"), theta1=modbus_get_signal_status("MiR_Theta_1"), theta2=modbus_get_signal_status("MiR_Theta_2"))
    $ 1167 "If MiR_Mode≠7"
    if (modbus_get_signal_status("MiR_Mode") != 7):
      $ 1168 "Error"
      $ 1169 "set_error(ERROR_AMR_WRONG_MODE)"
      set_error(ERROR_AMR_WRONG_MODE)
      $ 1170 "AMR_Done≔ True "
      global AMR_Done=  True
    end
    $ 1171 "'=========='"
    # '=========='
    $ 1172 "Switch STATE"
    switch_1 = STATE
    $ 1173 "Case 1"
    if (1 == switch_1):
      $ 1174 "stopping"
      $ 1175 "If T2O_Done≟1 and O2T_Acknowledge≟0"
      if (modbus_get_signal_status("T2O_Done") == 1  and  modbus_get_signal_status("O2T_Acknowledge") == 0):
        $ 1176 "Set O2T_Acknowledge=1"
        modbus_set_output_register("O2T_Acknowledge", 1)
      end
      $ 1177 "Set MiR_CMD_Stop=On"
      modbus_set_output_signal("MiR_CMD_Stop", True)
      $ 1178 "AMR_Position.position_identifier = 0"
      AMR_Position.position_identifier = 0
      $ 1179 "AMR_Done≔ True "
      global AMR_Done=  True
    elif (2 == switch_1):
      $ 1180 "Case 2"
      $ 1181 "stopped"
      $ 1182 "If MiR_State≠3 and MiR_State≠5"
      if (modbus_get_signal_status("MiR_State") != 3  and  modbus_get_signal_status("MiR_State") != 5):
        $ 1183 "Set MiR_CMD_Stop=Off"
        modbus_set_output_signal("MiR_CMD_Stop", False)
      end
    elif (3 == switch_1):
      $ 1184 "Case 3"
      $ 1185 "resetting"
      $ 1186 "Set O2T_Mis_Main=Off"
      modbus_set_output_signal("O2T_Mis_Main", False)
      $ 1187 "Set O2T_Mis_Charge=Off"
      modbus_set_output_signal("O2T_Mis_Charge", False)
      $ 1188 "If MiR_Mis_Queue>0"
      if (modbus_get_signal_status("MiR_Mis_Queue")>0):
        $ 1189 "Set MiR_CMD_Clear_Q=On"
        modbus_set_output_signal("MiR_CMD_Clear_Q", True)
        $ 1190 "Wait MiR_Mis_Queue≟0"
        while (not(modbus_get_signal_status("MiR_Mis_Queue") == 0)):
          sync()
        end
        $ 1191 "Set MiR_CMD_Clear_Q=Off"
        modbus_set_output_signal("MiR_CMD_Clear_Q", False)
      end
      $ 1192 "If MiR_Error_ID≠0"
      if (modbus_get_signal_status("MiR_Error_ID") != 0):
        $ 1193 "Set MiR_CMD_Clear_E=On"
        modbus_set_output_signal("MiR_CMD_Clear_E", True)
        $ 1194 "Wait MiR_Error_ID≟0"
        while (not(modbus_get_signal_status("MiR_Error_ID") == 0)):
          sync()
        end
        $ 1195 "Set MiR_CMD_Clear_E=Off"
        modbus_set_output_signal("MiR_CMD_Clear_E", False)
      end
      $ 1196 "Set O2T_Action=0"
      modbus_set_output_register("O2T_Action", 0)
      $ 1197 "Set O2T_Acknowledge=0"
      modbus_set_output_register("O2T_Acknowledge", 0)
      $ 1198 "Set O2T_Target_Pos=0"
      modbus_set_output_register("O2T_Target_Pos", 0)
      $ 1199 "Set O2T_Footprint=0"
      modbus_set_output_register("O2T_Footprint", 0)
      $ 1200 "Set O2T_ProtectOff=0"
      modbus_set_output_register("O2T_ProtectOff", 0)
      $ 1201 "Set O2T_Dock=0"
      modbus_set_output_register("O2T_Dock", 0)
      $ 1202 "AMR_Attemps≔0"
      global AMR_Attemps=0
      $ 1203 "AMR_PosTarget≔0"
      global AMR_PosTarget=0
      $ 1204 "AMR_Step≔0"
      global AMR_Step=0
      $ 1205 "AMR_AtTarget≔ False "
      global AMR_AtTarget=  False
      $ 1206 "If MiR_State≟4 or MiR_State≟3 or MiR_State≟10"
      if (modbus_get_signal_status("MiR_State") == 4  or  modbus_get_signal_status("MiR_State") == 3  or  modbus_get_signal_status("MiR_State") == 10):
        $ 1207 "AMR_Done≔ True "
        global AMR_Done=  True
      end
    elif (5 == switch_1):
      $ 1208 "Case 5"
      $ 1209 "starting"
      $ 1210 "If MiR_State≟4"
      if (modbus_get_signal_status("MiR_State") == 4):
        $ 1211 "Set MiR_CMD_Start=On"
        modbus_set_output_signal("MiR_CMD_Start", True)
        $ 1212 "Wait MiR_State≠4"
        while (not(modbus_get_signal_status("MiR_State") != 4)):
          sync()
        end
        $ 1213 "Set MiR_CMD_Start=Off"
        modbus_set_output_signal("MiR_CMD_Start", False)
        $ 1214 "AMR_Done≔ True "
        global AMR_Done=  True
      else:
        $ 1215 "ElseIf MiR_State≟10"
        if (modbus_get_signal_status("MiR_State") == 10):
          $ 1216 "'MiR in protective stop. Wait'"
          # 'MiR in protective stop. Wait'
          $ 1217 "AMR_Done≔ True "
          global AMR_Done=  True
        else:
          $ 1218 "ElseIf MiR_State≟3"
          if (modbus_get_signal_status("MiR_State") == 3):
            $ 1219 "AMR_Done≔ True "
            global AMR_Done=  True
          end
        end
      end
    elif (6 == switch_1):
      $ 1220 "Case 6"
      $ 1221 "execute"
      $ 1222 "AMR_AtTarget≔(AMR_PosActual≟AMR_PosTarget)"
      global AMR_AtTarget=(AMR_PosActual == AMR_PosTarget)
      $ 1223 "Switch AMR_Step"
      switch_2 = AMR_Step
      $ 1224 "Case 0"
      if (0 == switch_2):
        $ 1225 "If  not AMR_AtTarget"
        if (  not  AMR_AtTarget):
          $ 1226 "AMR_Step≔1"
          global AMR_Step=1
        else:
          $ 1227 "Else" "noBreak"
          $ 1228 "AMR_Done≔ True "
          global AMR_Done=  True
        end
      elif (1 == switch_2):
        $ 1229 "Case 1"
        $ 1230 "general Settings"
        $ 1231 "Set O2T_Acknowledge=0"
        modbus_set_output_register("O2T_Acknowledge", 0)
        $ 1232 "check for error"
        $ 1233 "If OBJ_Picked and MiR_State≟10"
        if (OBJ_Picked  and  modbus_get_signal_status("MiR_State") == 10):
          $ 1234 "Error"
          $ 1235 "set_error(ERROR_ROBOT_ARM_NOT_IN_HOME_POSE)"
          set_error(ERROR_ROBOT_ARM_NOT_IN_HOME_POSE)
          $ 1236 "Action≔0"
          global Action=0
        else:
          $ 1237 "ElseIf  not found_in_list(AMR_PosTarget, AMR_TargetList)"
          if (  not  found_in_list(AMR_PosTarget, AMR_TargetList)):
            $ 1238 "Error"
            $ 1239 "set_error(ERROR_UNKNOWN_POSE)"
            set_error(ERROR_UNKNOWN_POSE)
            $ 1240 "Action≔0"
            global Action=0
          end
        end
        $ 1241 "If MiR_State≟3"
        if (modbus_get_signal_status("MiR_State") == 3):
          $ 1242 "Set MiR_CMD_Start=Off"
          modbus_set_output_signal("MiR_CMD_Start", False)
          $ 1243 "Switch Action"
          switch_3 = Action
          $ 1244 "Case 51"
          if (51 == switch_3):
            $ 1245 "Charge"
            $ 1246 "'trigger the charging mission'"
            # 'trigger the charging mission'
            $ 1247 "'target pos is predefined'"
            # 'target pos is predefined'
            $ 1248 "Set O2T_Footprint=0"
            modbus_set_output_register("O2T_Footprint", 0)
            $ 1249 "Set O2T_Action=1"
            modbus_set_output_register("O2T_Action", 1)
            $ 1250 "If MiR_Mis_Queue≟0"
            if (modbus_get_signal_status("MiR_Mis_Queue") == 0):
              $ 1251 "Set O2T_Mis_Charge=On"
              modbus_set_output_signal("O2T_Mis_Charge", True)
              $ 1252 "Wait MiR_Mis_Queue≥1"
              while (not(modbus_get_signal_status("MiR_Mis_Queue") >= 1)):
                sync()
              end
              $ 1253 "Set O2T_Mis_Charge=Off"
              modbus_set_output_signal("O2T_Mis_Charge", False)
            end
          elif (52 == switch_3):
            $ 1254 "Case 52"
            $ 1255 "Navigate"
            $ 1256 "'trigger the standard missoin'"
            # 'trigger the standard missoin'
            $ 1257 "Set O2T_Footprint=AMR_FootprintID"
            modbus_set_output_register("O2T_Footprint", AMR_FootprintID)
            $ 1258 "Set O2T_Target_Pos=AMR_PosTarget"
            modbus_set_output_register("O2T_Target_Pos", AMR_PosTarget)
            $ 1259 "Set O2T_Action=2"
            modbus_set_output_register("O2T_Action", 2)
            $ 1260 "If MiR_Mis_Queue≟0"
            if (modbus_get_signal_status("MiR_Mis_Queue") == 0):
              $ 1261 "Set O2T_Mis_Main=On"
              modbus_set_output_signal("O2T_Mis_Main", True)
              $ 1262 "Wait MiR_Mis_Queue≥1"
              while (not(modbus_get_signal_status("MiR_Mis_Queue") >= 1)):
                sync()
              end
              $ 1263 "Set O2T_Mis_Main=Off"
              modbus_set_output_signal("O2T_Mis_Main", False)
            end
          end
        else:
          $ 1264 "ElseIf MiR_State≟4"
          if (modbus_get_signal_status("MiR_State") == 4):
            $ 1265 "Set MiR_CMD_Start=On"
            modbus_set_output_signal("MiR_CMD_Start", True)
          else:
            $ 1266 "ElseIf MiR_State≟5"
            if (modbus_get_signal_status("MiR_State") == 5):
              $ 1267 "AMR_Step≔2"
              global AMR_Step=2
            else:
              $ 1268 "ElseIf MiR_State≟10"
              if (modbus_get_signal_status("MiR_State") == 10):
                $ 1269 "'AMR still in safeguard stop'"
                # 'AMR still in safeguard stop'
              end
            end
          end
        end
      elif (2 == switch_2):
        $ 1270 "Case 2"
        $ 1271 "acknowledge handshake"
        $ 1272 "If T2O_Done≟1 and O2T_Acknowledge≟0"
        if (modbus_get_signal_status("T2O_Done") == 1  and  modbus_get_signal_status("O2T_Acknowledge") == 0):
          $ 1273 "Set O2T_Acknowledge=1"
          modbus_set_output_register("O2T_Acknowledge", 1)
        else:
          $ 1274 "ElseIf T2O_Done≟0 and O2T_Acknowledge≟1"
          if (modbus_get_signal_status("T2O_Done") == 0  and  modbus_get_signal_status("O2T_Acknowledge") == 1):
            $ 1275 "Set O2T_Acknowledge=0"
            modbus_set_output_register("O2T_Acknowledge", 0)
            $ 1276 "AMR_AtTarget≔(AMR_PosActual≟AMR_PosTarget)"
            global AMR_AtTarget=(AMR_PosActual == AMR_PosTarget)
            $ 1277 "AMR_Done≔ True "
            global AMR_Done=  True
          end
        end
      end
      $ 1278 "translate errors"
      $ 1279 "If AMR_Done"
      if (AMR_Done):
        $ 1280 "Switch T2O_Error_ID"
        switch_2 = modbus_get_signal_status("T2O_Error_ID")
        $ 1281 "Case 2003"
        if (2003 == switch_2):
          $ 1282 "error"
          $ 1283 "set_error(ERROR_NOT_DOCKED)"
          set_error(ERROR_NOT_DOCKED)
        elif (2007 == switch_2):
          $ 1284 "Case 2007"
          $ 1285 "error"
          $ 1286 "set_error(ERROR_NOT_REACHABLE_TARGET)"
          set_error(ERROR_NOT_REACHABLE_TARGET)
        elif (2008 == switch_2):
          $ 1287 "Case 2008"
          $ 1288 "error"
          $ 1289 "set_error(ERROR_CHARGING_NOT_STARTED)"
          set_error(ERROR_CHARGING_NOT_STARTED)
        end
      end
    elif (7 == switch_1):
      $ 1290 "Case 7"
      $ 1291 "completing"
      $ 1292 "If MiR_Mis_Queue>0"
      if (modbus_get_signal_status("MiR_Mis_Queue")>0):
        $ 1293 "Set MiR_CMD_Abort=On"
        modbus_set_output_signal("MiR_CMD_Abort", True)
        $ 1294 "Wait MiR_Mis_Queue≟0"
        while (not(modbus_get_signal_status("MiR_Mis_Queue") == 0)):
          sync()
        end
        $ 1295 "Set MiR_CMD_Abort=Off"
        modbus_set_output_signal("MiR_CMD_Abort", False)
      end
      $ 1296 "If MiR_State≟3 or MiR_State≟10"
      if (modbus_get_signal_status("MiR_State") == 3  or  modbus_get_signal_status("MiR_State") == 10):
        $ 1297 "AMR_Done≔ True "
        global AMR_Done=  True
      end
    elif (9 == switch_1):
      $ 1298 "Case 9"
      $ 1299 "holding"
      $ 1300 "Set MiR_CMD_Abort=On"
      modbus_set_output_signal("MiR_CMD_Abort", True)
      $ 1301 "If MiR_State≟3 or MiR_State≟10"
      if (modbus_get_signal_status("MiR_State") == 3  or  modbus_get_signal_status("MiR_State") == 10):
        $ 1302 "Set MiR_CMD_Abort=Off"
        modbus_set_output_signal("MiR_CMD_Abort", False)
        $ 1303 "AMR_Done≔ True "
        global AMR_Done=  True
      end
    elif (11 == switch_1):
      $ 1304 "Case 11"
      $ 1305 "unholding"
      $ 1306 "Set MiR_CMD_Start=On"
      modbus_set_output_signal("MiR_CMD_Start", True)
      $ 1307 "If MiR_State≠4"
      if (modbus_get_signal_status("MiR_State") != 4):
        $ 1308 "Set MiR_CMD_Start=Off"
        modbus_set_output_signal("MiR_CMD_Start", False)
        $ 1309 "AMR_Step≔0"
        global AMR_Step=0
        $ 1310 "AMR_Done≔ True "
        global AMR_Done=  True
      end
    elif (12 == switch_1):
      $ 1311 "Case 12"
      $ 1312 "suspending"
      $ 1313 "'none'"
      # 'none'
    elif (14 == switch_1):
      $ 1314 "Case 14"
      $ 1315 "unsuspending"
      $ 1316 "'none'"
      # 'none'
    elif (15 == switch_1):
      $ 1317 "Case 15"
      $ 1318 "aborting"
      $ 1319 "Set MiR_CMD_Abort=On"
      modbus_set_output_signal("MiR_CMD_Abort", True)
      $ 1320 "Wait MiR_State≟3"
      while (not(modbus_get_signal_status("MiR_State") == 3)):
        sync()
      end
      $ 1321 "Set MiR_CMD_Abort=Off"
      modbus_set_output_signal("MiR_CMD_Abort", False)
    elif (17 == switch_1):
      $ 1322 "Case 17"
      $ 1323 "clearing"
      $ 1324 "If MiR_Error_ID≠0"
      if (modbus_get_signal_status("MiR_Error_ID") != 0):
        $ 1325 "Set MiR_CMD_Clear_E=On"
        modbus_set_output_signal("MiR_CMD_Clear_E", True)
        $ 1326 "Wait MiR_Error_ID≟0"
        while (not(modbus_get_signal_status("MiR_Error_ID") == 0)):
          sync()
        end
        $ 1327 "Set MiR_CMD_Clear_E=Off"
        modbus_set_output_signal("MiR_CMD_Clear_E", False)
      end
      $ 1328 "If MiR_Error_ID≟0"
      if (modbus_get_signal_status("MiR_Error_ID") == 0):
        $ 1329 "AMR_Done≔ True "
        global AMR_Done=  True
      end
    end
    $ 1330 "'=========='"
    # '=========='
    $ 1331 "PostSettings"
    $ 1332 "AMR_Position≔struct(position_identifier=T2O_Current_Pos, x1=MiR_Position_X1, x2=MiR_Position_X2, y1=MiR_Position_Y1, y2=MiR_Position_Y2, theta1=MiR_Theta_1, theta2=MiR_Theta_2) "
    global AMR_Position=struct(position_identifier=modbus_get_signal_status("T2O_Current_Pos"), x1=modbus_get_signal_status("MiR_Position_X1"), x2=modbus_get_signal_status("MiR_Position_X2"), y1=modbus_get_signal_status("MiR_Position_Y1"), y2=modbus_get_signal_status("MiR_Position_Y2"), theta1=modbus_get_signal_status("MiR_Theta_1"), theta2=modbus_get_signal_status("MiR_Theta_2"))
  end
  def Sub_Action_V4():
    $ 1333 "Sub_Action_V4" "noBreak"
    $ 1334 "PreSettings"
    $ 1335 "init poses"
    $ 1336 "PSE_A≔p[0,0,0,0,0,0]"
    global PSE_A=p[0,0,0,0,0,0]
    $ 1337 "PSE_A_H≔p[0,0,0,0,0,0]"
    global PSE_A_H=p[0,0,0,0,0,0]
    $ 1338 "PSE_T≔p[0,0,0,0,0,0]"
    global PSE_T=p[0,0,0,0,0,0]
    $ 1339 "PSE_T_H≔p[0,0,0,0,0,0]"
    global PSE_T_H=p[0,0,0,0,0,0]
    $ 1340 "PSE_G≔p[0,0,0,0,0,0]"
    global PSE_G=p[0,0,0,0,0,0]
    $ 1341 "PSE_G_H≔p[0,0,0,0,0,0]"
    global PSE_G_H=p[0,0,0,0,0,0]
    $ 1342 "PSE_R≔p[0,0,0,0,0,0]"
    global PSE_R=p[0,0,0,0,0,0]
    $ 1343 "PSE_R_H≔p[0,0,0,0,0,0]"
    global PSE_R_H=p[0,0,0,0,0,0]
    $ 1344 "JNT_Q≔[0,0,0,0,0,0]"
    global JNT_Q=[0,0,0,0,0,0]
    $ 1345 "JNT_S≔[0,0,0,0,0,0]"
    global JNT_S=[0,0,0,0,0,0]
    $ 1346 "Gripping parameters"
    $ 1347 "OBJ = find_object_by_type(OBJs, OBJ_Type)"
    OBJ = find_object_by_type(OBJs, OBJ_Type)
    $ 1348 "GRP_Open_Pos≔OBJ.dimension.diameter * 1000 + 6"
    global GRP_Open_Pos=OBJ.dimension.diameter * 1000 + 6
    $ 1349 "GRP_Offset≔OBJ.gripper_offset"
    global GRP_Offset=OBJ.gripper_offset
    $ 1350 "rq_set_force_norm(50)"
     rq_set_force_norm (50)
    $ 1351 "rq_set_speed_norm(50)"
     rq_set_speed_norm (50)
    $ 1352 "Switch ITM_ID"
    switch_1 = ITM_ID
    $ 1353 "Case 1"
    if (1 == switch_1):
      $ 1354 "uML"
      $ 1355 "JIG2 = find_object_by_type(JIGs, JIG)"
      JIG2 = find_object_by_type(JIGs, JIG)
      $ 1356 "JIG_Offset≔JIG2.jig_offset"
      global JIG_Offset=JIG2.jig_offset
      $ 1357 "Switch JIG"
      switch_2 = JIG
      $ 1358 "Case 1"
      if (1 == switch_2):
        $ 1359 "3FG"
        $ 1360 "define poses"
        $ 1361 "FRM_Reference≔ULM_3FG"
        global FRM_Reference=ULM_3FG
        $ 1362 "JNT_Q≔JNT_HOME"
        global JNT_Q=JNT_HOME
        $ 1363 "PSE_T≔pose_trans(GRP_Offset, JIG_Offset)"
        global PSE_T= pose_trans (GRP_Offset, JIG_Offset)
        $ 1364 "PSE_A≔pose_trans(PSE_T, p[0,0,0.100,0,0,0])"
        global PSE_A= pose_trans (PSE_T, p[0,0,0.100,0,0,0])
        $ 1365 "PSE_R≔pose_add(PSE_T, p[0,0,0.100,0,0,0])"
        global PSE_R= pose_add (PSE_T, p[0,0,0.100,0,0,0])
      elif (2 == switch_2):
        $ 1366 "Case 2"
        $ 1367 "Input"
        $ 1368 "'CHANGE THE REFERENCE TO THE FRAME TO MOVE IN'"
        # 'CHANGE THE REFERENCE TO THE FRAME TO MOVE IN'
        $ 1369 "define poses"
        $ 1370 "FRM_Reference≔ULM_Input"
        global FRM_Reference=ULM_Input
        $ 1371 "PSE_T≔pose_trans(pose_trans(get_pattern_pos_rectangle(OBJ_Nbr, 'X', [10,5], patternsize=[0.181,0.081]), GRP_Offset), JIG_Offset)"
        global PSE_T= pose_trans ( pose_trans (get_pattern_pos_rectangle(OBJ_Nbr, "X", [10,5], patternsize=[0.181,0.081]), GRP_Offset), JIG_Offset)
        $ 1372 "If Action≟1"
        if (Action == 1):
          $ 1373 "PSE_R≔pose_add(PSE_T, p[0,0,0.200,0,0,0])"
          global PSE_R= pose_add (PSE_T, p[0,0,0.200,0,0,0])
          $ 1374 "PSE_A≔pose_add(PSE_T, p[0,0,0.100,0,0,0])"
          global PSE_A= pose_add (PSE_T, p[0,0,0.100,0,0,0])
        else:
          $ 1375 "ElseIf Action≟2"
          if (Action == 2):
            $ 1376 "PSE_R≔pose_add(PSE_T, p[0,0,0.100,0,0,0])"
            global PSE_R= pose_add (PSE_T, p[0,0,0.100,0,0,0])
            $ 1377 "PSE_A≔pose_add(PSE_T, p[0,0,0.200,0,0,0])"
            global PSE_A= pose_add (PSE_T, p[0,0,0.200,0,0,0])
          end
        end
      elif (3 == switch_2):
        $ 1378 "Case 3"
        $ 1379 "Output"
        $ 1380 "'CHANGE THE REFERENCE TO THE FRAME TO MOVE IN'"
        # 'CHANGE THE REFERENCE TO THE FRAME TO MOVE IN'
        $ 1381 "define poses"
        $ 1382 "FRM_Reference≔ULM_Output"
        global FRM_Reference=ULM_Output
        $ 1383 "PSE_T≔pose_trans(pose_trans(get_pattern_pos_rectangle(OBJ_Nbr, 'X', [10,5], patternsize=[0.181,0.081]), GRP_Offset), JIG_Offset)"
        global PSE_T= pose_trans ( pose_trans (get_pattern_pos_rectangle(OBJ_Nbr, "X", [10,5], patternsize=[0.181,0.081]), GRP_Offset), JIG_Offset)
        $ 1385 "If Action≟1"
        if (Action == 1):
          $ 1386 "PSE_R≔pose_add(PSE_T, p[0,0,0.200,0,0,0])"
          global PSE_R= pose_add (PSE_T, p[0,0,0.200,0,0,0])
          $ 1387 "PSE_A≔pose_add(PSE_T, p[0,0,0.100,0,0,0])"
          global PSE_A= pose_add (PSE_T, p[0,0,0.100,0,0,0])
        else:
          $ 1388 "ElseIf Action≟2"
          if (Action == 2):
            $ 1389 "PSE_R≔pose_add(PSE_T, p[0,0,0.100,0,0,0])"
            global PSE_R= pose_add (PSE_T, p[0,0,0.100,0,0,0])
            $ 1390 "PSE_A≔pose_add(PSE_T, p[0,0,0.200,0,0,0])"
            global PSE_A= pose_add (PSE_T, p[0,0,0.200,0,0,0])
          end
        end
      elif (4 == switch_2):
        $ 1391 "Case 4"
        $ 1392 "jig centrifuge racks"
        $ 1393 "define poses"
        $ 1394 "FRM_Reference≔ULM_Cent_Racks"
        global FRM_Reference=ULM_Cent_Racks
        $ 1395 "PSE_T≔get_pattern_pos_rectangle(JIG_Slot, 'X', [4,1], patternsize=[0.291,0])"
        global PSE_T=get_pattern_pos_rectangle(JIG_Slot, "X", [4,1], patternsize=[0.291,0])
        $ 1396 "If OBJ_Nbr≠0"
        if (OBJ_Nbr != 0):
          $ 1397 "PSE_T≔pose_trans(pose_trans(PSE_T, get_pattern_pos_rectangle(OBJ_Nbr, 'X', [3,3], patternsize=[0.060,0.060])),p[-0.030, -0.030,0,0,0,3.927])"
          global PSE_T= pose_trans ( pose_trans (PSE_T, get_pattern_pos_rectangle(OBJ_Nbr, "X", [3,3], patternsize=[0.060,0.060])),p[-0.030, -0.030,0,0,0,3.927])
        end
        $ 1398 "PSE_T≔pose_trans(PSE_T, GRP_Offset)"
        global PSE_T= pose_trans (PSE_T, GRP_Offset)
        $ 1399 "If Action≟1"
        if (Action == 1):
          $ 1400 "PSE_R≔pose_add(PSE_T, p[0,0,0.200,0,0,0])"
          global PSE_R= pose_add (PSE_T, p[0,0,0.200,0,0,0])
          $ 1401 "PSE_A≔pose_add(PSE_T, p[0,0,0.100,0,0,0])"
          global PSE_A= pose_add (PSE_T, p[0,0,0.100,0,0,0])
        else:
          $ 1402 "ElseIf Action≟2"
          if (Action == 2):
            $ 1403 "PSE_R≔pose_add(PSE_T, p[0,0,0.100,0,0,0])"
            global PSE_R= pose_add (PSE_T, p[0,0,0.100,0,0,0])
            $ 1404 "PSE_A≔pose_add(PSE_T, p[0,0,0.200,0,0,0])"
            global PSE_A= pose_add (PSE_T, p[0,0,0.200,0,0,0])
          end
        end
      elif (6 == switch_2):
        $ 1405 "Case 6"
        $ 1406 "Caps bin"
        $ 1407 "define poses"
        $ 1408 "'Drop cap'"
        # 'Drop cap'
        $ 1409 "FRM_Reference=ULM_Cap_Bin"
        FRM_Reference=ULM_Cap_Bin
        $ 1410 "PSE_T≔pose_RPY2RotVec(p[0,0,0,0,0,0])"
        global PSE_T=pose_RPY2RotVec(p[0,0,0,0,0,0])
        $ 1411 "PSE_T_H≔pose_add(PSE_T, p[0,0,-0.011,0,0,0])"
        global PSE_T_H= pose_add (PSE_T, p[0,0,-0.011,0,0,0])
        $ 1412 "PSE_A≔pose_trans(PSE_T, p[0,0,0.1,0,0,0])"
        global PSE_A= pose_trans (PSE_T, p[0,0,0.1,0,0,0])
        $ 1413 "PSE_R_H≔pose_add(PSE_T, p[0,0,0.100,0,0,0])"
        global PSE_R_H= pose_add (PSE_T, p[0,0,0.100,0,0,0])
        $ 1414 "PSE_R≔pose_add(PSE_T, p[0,0,0.100,0,0,0])"
        global PSE_R= pose_add (PSE_T, p[0,0,0.100,0,0,0])
      elif (7 == switch_2):
        $ 1415 "Case 7"
        $ 1416 "Sarstedt"
        $ 1417 "'CHANGE THE REFERENCE TO THE FRAME TO MOVE IN'"
        # 'CHANGE THE REFERENCE TO THE FRAME TO MOVE IN'
        $ 1423 "If TASK.ID≟10"
        if (TASK.ID == 10):
          $ 1424 "Frame & Position Params"
          $ 1426 "FRM_Reference = CAM_LM_SSRack"
          FRM_Reference = CAM_LM_SSRack
          $ 1431 "PSE_T≔uLM_SS_PickPlc"
          global PSE_T=uLM_SS_PickPlc
          $ 1432 "PSE_A≔pose_trans(PSE_T, p[0,0,0.1,0,0,0])"
          global PSE_A= pose_trans (PSE_T, p[0,0,0.1,0,0,0])
          $ 1433 "PSE_R≔pose_add(PSE_T, p[0,0,0.1,0,0,0])"
          global PSE_R= pose_add (PSE_T, p[0,0,0.1,0,0,0])
        else:
          $ 1434 "ElseIf TASK.ID≟11"
          if (TASK.ID == 11):
            $ 1435 "FRM_Reference = ULM_SS_Jig"
            FRM_Reference = ULM_SS_Jig
            $ 1436 "PSE_T≔pose_RPY2RotVec(p[0,0,0,0,0,0])"
            global PSE_T=pose_RPY2RotVec(p[0,0,0,0,0,0])
            $ 1437 "PSE_T≔pose_trans(PSE_T, GRP_Offset)"
            global PSE_T=pose_trans(PSE_T, GRP_Offset)
            $ 1438 "PSE_A≔pose_trans(PSE_T, p[0,0,0.1,0,0,0])"
            global PSE_A= pose_trans (PSE_T, p[0,0,0.1,0,0,0])
            $ 1439 "PSE_R≔pose_add(PSE_T, p[0,0,0.2,0,0,0])"
            global PSE_R= pose_add (PSE_T, p[0,0,0.2,0,0,0])
          end
        end
      elif (8 == switch_2):
        $ 1440 "Case 8"
        $ 1441 "NoK"
        $ 1442 "define poses"
        $ 1443 "'NoK'"
        # 'NoK'
        $ 1444 "FRM_Reference=ULM_NoK"
        FRM_Reference=ULM_NoK
        $ 1445 "PSE_T≔pose_RPY2RotVec(p[0,0,0,0,0,0])"
        global PSE_T=pose_RPY2RotVec(p[0,0,0,0,0,0])
        $ 1446 "PSE_A≔pose_trans(PSE_T, p[0,0,0.1,0,0,0])"
        global PSE_A= pose_trans (PSE_T, p[0,0,0.1,0,0,0])
        $ 1447 "PSE_R≔pose_add(PSE_T, p[0,0,0.100,0,0,0])"
        global PSE_R= pose_add (PSE_T, p[0,0,0.100,0,0,0])
      elif (9 == switch_2):
        $ 1448 "Case 9"
        $ 1449 "Pick_bott_jig"
        $ 1450 "define poses"
        $ 1451 "'NoK'"
        # 'NoK'
        $ 1452 "FRM_Reference=ULM_bottle_pick_const"
        FRM_Reference=p[0.08175869478771049,-0.47602162643540935,0.09,0.00141829700319658,-0.0027789445191063835,0.07763675748118615]
        $ 1453 "PSE_T≔pose_RPY2RotVec(p[0,0,0,0,0,0])"
        global PSE_T=pose_RPY2RotVec(p[0,0,0,0,0,0])
        $ 1454 "PSE_A≔pose_trans(PSE_T, p[0,0,0.1,0,0,0])"
        global PSE_A= pose_trans (PSE_T, p[0,0,0.1,0,0,0])
        $ 1455 "PSE_R≔pose_add(PSE_T, p[0,0,0.100,0,0,0])"
        global PSE_R= pose_add (PSE_T, p[0,0,0.100,0,0,0])
      elif (10 == switch_2):
        $ 1456 "Case 10"
        $ 1457 "Place_bott_jig"
        $ 1458 "define poses"
        $ 1459 "'NoK'"
        # 'NoK'
        $ 1460 "FRM_Reference=ULM_bottle_plac_const"
        FRM_Reference=p[-0.09502738395762109,-0.5154087721098056,0.095,0.0014590126708889871,-0.0028280855286173575,0.07763149296298452]
        $ 1461 "PSE_T≔pose_RPY2RotVec(p[0,0,0,0,0,0])"
        global PSE_T=pose_RPY2RotVec(p[0,0,0,0,0,0])
        $ 1462 "PSE_A≔pose_trans(PSE_T, p[0,0,0.1,0,0,0])"
        global PSE_A= pose_trans (PSE_T, p[0,0,0.1,0,0,0])
        $ 1463 "PSE_R≔pose_add(PSE_T, p[0,0,0.100,0,0,0])"
        global PSE_R= pose_add (PSE_T, p[0,0,0.100,0,0,0])
      elif (11 == switch_2):
        $ 1464 "Case 11"
        $ 1465 "Place_bott_jig"
        $ 1466 "define poses"
        $ 1467 "'NoK'"
        # 'NoK'
        $ 1468 "FRM_Reference=shake"
        FRM_Reference=shake
        $ 1469 "PSE_T≔pose_RPY2RotVec(p[0,0,0,0,0,0])"
        global PSE_T=pose_RPY2RotVec(p[0,0,0,0,0,0])
        $ 1470 "PSE_A≔pose_trans(PSE_T, p[0,0,0,0,0,0])"
        global PSE_A= pose_trans (PSE_T, p[0,0,0,0,0,0])
        $ 1471 "PSE_R≔pose_add(PSE_T, p[0,0,0,0,0,0])"
        global PSE_R= pose_add (PSE_T, p[0,0,0,0,0,0])
      elif (12 == switch_2):
        $ 1472 "Case 12"
        $ 1473 "Pick_Vial_jig"
        $ 1474 "define poses"
        $ 1475 "'NoK'"
        # 'NoK'
        $ 1476 "FRM_Reference=shake"
        FRM_Reference=shake
        $ 1477 "PSE_T≔pose_RPY2RotVec(p[0,0,0,0,0,0])"
        global PSE_T=pose_RPY2RotVec(p[0,0,0,0,0,0])
        $ 1478 "PSE_A≔pose_trans(PSE_T, p[0,0,0,0,0,0])"
        global PSE_A= pose_trans (PSE_T, p[0,0,0,0,0,0])
        $ 1479 "PSE_R≔pose_add(PSE_T, p[0,0,0,0,0,0])"
        global PSE_R= pose_add (PSE_T, p[0,0,0,0,0,0])
      end
    elif (2 == switch_1):
      $ 1480 "Case 2"
      $ 1481 "Centrifuge"
      $ 1482 "'CHANGE THE REFERENCE TO THE FRAME TO MOVE IN'"
      # 'CHANGE THE REFERENCE TO THE FRAME TO MOVE IN'
      $ 1483 "define poses"
      $ 1484 "FRM_Reference≔FRM_Centrifuge"
      global FRM_Reference=FRM_Centrifuge
      $ 1485 "PSE_T≔GRP_Offset"
      global PSE_T=GRP_Offset
      $ 1486 "If Action≟8"
      if (Action == 8):
        $ 1487 "PSE_R≔pose_add(PSE_T, p[0,0,0.250,0,0,0])"
        global PSE_R= pose_add (PSE_T, p[0,0,0.250,0,0,0])
        $ 1488 "PSE_A≔pose_add(PSE_T, p[0,0,0.150,0,0,0])"
        global PSE_A= pose_add (PSE_T, p[0,0,0.150,0,0,0])
      else:
        $ 1489 "ElseIf Action≟7"
        if (Action == 7):
          $ 1490 "PSE_R≔pose_add(PSE_T, p[0,0,0.150,0,0,0])"
          global PSE_R= pose_add (PSE_T, p[0,0,0.150,0,0,0])
          $ 1491 "PSE_A≔pose_add(PSE_T, p[0,0,0.250,0,0,0])"
          global PSE_A= pose_add (PSE_T, p[0,0,0.250,0,0,0])
        end
      end
    elif (3 == switch_1):
      $ 1492 "Case 3"
      $ 1493 "Output"
      $ 1494 "'CHANGE THE REFERENCE TO THE FRAME TO MOVE IN'"
      # 'CHANGE THE REFERENCE TO THE FRAME TO MOVE IN'
      $ 1495 "define poses"
      $ 1496 "FRM_Reference≔Base_const"
      global FRM_Reference=p[0.0,0.0,0.0,0.0,0.0,0.0]
      $ 1497 "PSE_T≔p[0,0,0,0,0,0]"
      global PSE_T=p[0,0,0,0,0,0]
      $ 1498 "PSE_A≔pose_add(PSE_T, p[0,0,0.150,0,0,0])"
      global PSE_A= pose_add (PSE_T, p[0,0,0.150,0,0,0])
      $ 1499 "PSE_R≔pose_add(PSE_T, p[0,0,0.100,0,0,0])"
      global PSE_R= pose_add (PSE_T, p[0,0,0.100,0,0,0])
    elif (5 == switch_1):
      $ 1500 "Case 5"
      $ 1501 "Sarstedt Pickup Table"
      $ 1502 "'CHANGE THE REFERENCE TO THE FRAME TO MOVE IN'"
      # 'CHANGE THE REFERENCE TO THE FRAME TO MOVE IN'
      $ 1503 "Switch JIG"
      switch_2 = JIG
      $ 1504 "Case 7"
      if (7 == switch_2):
        $ 1517 "Sarstedt"
        $ 1518 "'CHANGE THE REFERENCE TO THE FRAME TO MOVE IN'"
        # 'CHANGE THE REFERENCE TO THE FRAME TO MOVE IN'
        $ 1524 "If TASK.ID≟10"
        if (TASK.ID == 10):
          $ 1525 "Frame & Position Params"
          $ 1526 "FRM_Reference = CAM_LM_SSRack"
          FRM_Reference = CAM_LM_SSRack
          $ 1527 "PSE_T≔uLM_SS_PickPlc"
          global PSE_T=uLM_SS_PickPlc
          $ 1528 "PSE_A≔pose_trans(PSE_T, p[0,0,0.1,0,0,0])"
          global PSE_A= pose_trans (PSE_T, p[0,0,0.1,0,0,0])
          $ 1529 "PSE_R≔pose_add(PSE_T, p[0,0,0.1,0,0,0])"
          global PSE_R= pose_add (PSE_T, p[0,0,0.1,0,0,0])
        end
      end
    elif (13 == switch_1):
      $ 1536 "Case 13"
      $ 1537 "Sarstedt Pickup Table"
      $ 1538 "'CHANGE THE REFERENCE TO THE FRAME TO MOVE IN'"
      # 'CHANGE THE REFERENCE TO THE FRAME TO MOVE IN'
      $ 1539 "Switch JIG"
      switch_2 = JIG
      $ 1540 "Case 7"
      if (7 == switch_2):
        $ 1553 "Bottle"
        $ 1554 "'CHANGE THE REFERENCE TO THE FRAME TO MOVE IN'"
        # 'CHANGE THE REFERENCE TO THE FRAME TO MOVE IN'
        $ 1560 "If TASK.ID≟43"
        if (TASK.ID == 43):
          $ 1561 "Frame & Position Params"
          $ 1562 "FRM_Reference = CAM_LM_Bott"
          FRM_Reference = CAM_LM_Bott
          $ 1563 "PSE_T≔uLM_SS_PickPlc"
          global PSE_T=uLM_SS_PickPlc
          $ 1564 "PSE_A≔pose_trans(PSE_T, p[0,0,0.1,0,0,0])"
          global PSE_A= pose_trans (PSE_T, p[0,0,0.1,0,0,0])
          $ 1565 "PSE_R≔pose_add(PSE_T, p[0,0,0.1,0,0,0])"
          global PSE_R= pose_add (PSE_T, p[0,0,0.1,0,0,0])
        end
      end
    end
    $ 1572 "Additional check"
    $ 1573 "If  not is_reachable(FRM_Reference,[PSE_A,PSE_A_H,PSE_T,PSE_T_H,PSE_R,PSE_R_H])"
    if (  not  is_reachable(FRM_Reference,[PSE_A,PSE_A_H,PSE_T,PSE_T_H,PSE_R,PSE_R_H])):
      $ 1574 "Error"
      $ 1575 "set_error(ERROR_POSE_NOT_REACHABLE)"
      set_error(ERROR_POSE_NOT_REACHABLE)
      $ 1576 "Action≔0"
      global Action=0
    end
    $ 1577 "'=========='"
    # '=========='
    $ 1578 "Switch Action"
    switch_1 = Action
    $ 1579 "Case 1"
    if (1 == switch_1):
      $ 1580 "Pick"
      $ 1581 "Action_Info≔'pick object'"
      global Action_Info="pick object"
      $ 1582 "do_transition(pose_trans(FRM_Reference, PSE_T), keep_rxry=OBJ_Picked)"
      do_transition( pose_trans (FRM_Reference, PSE_T), keep_rxry=OBJ_Picked)
      $ 1583 "EOAT"
      $ 1584 "If  not OBJ_Picked"
      if (  not  OBJ_Picked):
        $ 1585 "rq_move_and_wait_mm(GRP_Open_Pos)"
         rq_move_and_wait_mm (GRP_Open_Pos)
      end
      $ 1586 "If PSE_A_H≠PSE_Z"
      if (PSE_A_H != PSE_Z):
        $ 1587 "If JNT_Q≠JNT_Z"
        if (JNT_Q != JNT_Z):
          $ 1588 "movej(get_inverse_kin(pose_trans(FRM_Reference, PSE_A_H), qnear=JNT_Q), r=0.050)"
          movej(get_inverse_kin( pose_trans (FRM_Reference, PSE_A_H), qnear=JNT_Q), r=0.050)
        else:
          $ 1589 "Else" "noBreak"
          $ 1590 "movej(pose_trans(FRM_Reference, PSE_A_H), r=0.050)"
          movej( pose_trans (FRM_Reference, PSE_A_H), r=0.050)
        end
      end
      $ 1591 "If PSE_A≠PSE_Z"
      if (PSE_A != PSE_Z):
        $ 1592 "If JNT_Q≠JNT_Z"
        if (JNT_Q != JNT_Z):
          $ 1593 "movej(get_inverse_kin(pose_trans(FRM_Reference, PSE_A), qnear=JNT_Q), r=0.020)"
          movej(get_inverse_kin( pose_trans (FRM_Reference, PSE_A), qnear=JNT_Q), r=0.020)
        else:
          $ 1594 "Else" "noBreak"
          $ 1595 "movej(pose_trans(FRM_Reference, PSE_A), r=0.020)"
          movej( pose_trans (FRM_Reference, PSE_A), r=0.020)
        end
      end
      $ 1596 "MoveL"
      $ 1597 "If PSE_T_H≠PSE_Z"
      if (PSE_T_H != PSE_Z):
        $ 1598 "PSE_T_H" "breakAfter"
        movel(pose_trans(FRM_Reference, PSE_T_H), a=0.5, v=0.4, r=0.01)
      end
      $ 1599 "PSE_T" "breakAfter"
      movel(pose_trans(FRM_Reference, PSE_T), a=0.08, v=0.12)
      $ 1600 "EOAT"
      $ 1601 "rq_set_force_norm(50)"
       rq_set_force_norm (50)
      $ 1602 "rq_close_and_wait()"
       rq_close_and_wait ()
      $ 1603 "OBJ_Picked≔rq_is_object_detected()"
      global OBJ_Picked= rq_is_object_detected ()
      $ 1604 "If  not OBJ_Picked"
      if (  not  OBJ_Picked):
        $ 1605 "set_error(ERROR_NO_OBJECT_TO_PICK)"
        set_error(ERROR_NO_OBJECT_TO_PICK)
      end
      $ 1606 "EXTT"
      $ 1607 "Switch JIG"
      switch_2 = JIG
      $ 1608 "Case 1"
      if (1 == switch_2):
        $ 1609 "3FG"
        $ 1610 "If OBJ_Picked"
        if (OBJ_Picked):
          $ 1611 "Set GRP_3F_Open=On"
          set_standard_digital_out(5, True)
        end
      end
      $ 1612 "If PSE_R_H≠PSE_Z"
      if (PSE_R_H != PSE_Z):
        $ 1613 "PSE_R" "breakAfter"
        movel(pose_trans(FRM_Reference, PSE_R), a=0.5, v=0.4, r=0.01)
        $ 1614 "PSE_R_H" "breakAfter"
        movel(pose_trans(FRM_Reference, PSE_R_H), a=0.5, v=0.4)
      else:
        $ 1615 "Else" "noBreak"
        $ 1616 "PSE_R" "breakAfter"
        movel(pose_trans(FRM_Reference, PSE_R), a=0.5, v=0.4)
      end
    elif (2 == switch_1):
      $ 1617 "Case 2"
    elif (3 == switch_1):
      $ 1659 "Case 3"
    elif (4 == switch_1):
      $ 1662 "Case 4"
    elif (6 == switch_1):
      $ 1665 "Case 6"
    elif (7 == switch_1):
      $ 1680 "Case 7"
    elif (8 == switch_1):
      $ 1709 "Case 8"
    elif (11 == switch_1):
      $ 1742 "Case 11"
    elif (12 == switch_1):
      $ 1779 "Case 12"
    elif (15 == switch_1):
      $ 1830 "Case 15"
    elif (30 == switch_1):
      $ 1833 "Case 30"
    elif (31 == switch_1):
      $ 1866 "Case 31"
    elif (32 == switch_1):
      $ 1878 "Case 32"
    elif (33 == switch_1):
      $ 1919 "Case 33"
    elif (35 == switch_1):
      $ 1985 "Case 35"
      $ 1986 "Pick the powder container"
      # begin: URCap Program Node
      #   Source: SensoPart VISOR Robotic, 2.0.0, SensoPart Industriesensorik GmbH
      #   Type: VISOR Robotic App
      $ 1989 "VISOR Easy Pick"
      def visorFuncEasyPick_084428():
        # begin: URCap Program Node
        #   Source: SensoPart VISOR Robotic, 2.0.0, SensoPart Industriesensorik GmbH
        #   Type: Easy Pick Setup
        $ 1990 "# 1 Setup" "noBreak"
        local easyPickVisorId = 1
        local easyPickArmMounted = True
        local easyPickSetJob = True
        local easyPickJobName = "Container"
        local easyPickAtImgAcq = False
        local easyPickImgAcqPose = cont_img_pose
        # end: URCap Program Node
        # begin: URCap Program Node
        #   Source: SensoPart VISOR Robotic, 2.0.0, SensoPart Industriesensorik GmbH
        #   Type: Process
        $ 1991 "Process" "noBreak"
        local easyPickObjTaken = False
        local easyPickTrigger = False
        local easyPickPoseIdx = 0
        local easyPickPose = p[0,0,0,0,0,0]
        def easyPickFuncTrigger(visorId, setJob, jobName, arm):
        if (setJob):
          visor_changeJob(visorId, jobName, 6000)
        end
        if (arm):
          visor_trigger(visorId, 6000, "arm")
        else:
          visor_trigger(visorId, 6000)
        end
        global easyPickParts=visor_partsFound(visorId)
        visor_easyPickUpdate(visorId, "parts", visor_partsFound(visorId))
        return visor_getPose3d(visorId, 0)
      end
      while (not easyPickObjTaken):
        easyPickTrigger = (easyPickCount >= visor_partsFound(easyPickVisorId)) or (easyPickCount > 9) or (not visor_easyPickCheckIdent("9ca581", easyPickVisorId))
        if (easyPickTrigger):
          easyPickCount = 0
        end
        easyPickPoseIdx = easyPickCount
        easyPickPose = visor_getPose3d(easyPickVisorId, easyPickPoseIdx)
        visor_easyPickUpdate(easyPickVisorId, "counter", easyPickPoseIdx)
        # begin: URCap Program Node
        #   Source: SensoPart VISOR Robotic, 2.0.0, SensoPart Industriesensorik GmbH
        #   Type: Image Acquisition Pose
        $ 1992 "Image Acquisition Pose" "noBreak"
        if (easyPickTrigger):
          if (not easyPickAtImgAcq):
            movej(pose_trans(easyPickImgAcqPose,p[0.0000,0.0000,-0.0000,0.0000,0.0000,0.0000]),a=1.3963,v=1.0472,t=0.000000,r=0.000000)
            easyPickAtImgAcq = True
          end
          easyPickPose = easyPickFuncTrigger(easyPickVisorId, easyPickSetJob, easyPickJobName, easyPickArmMounted)
        end
        # end: URCap Program Node
        # begin: URCap Program Node
        #   Source: SensoPart VISOR Robotic, 2.0.0, SensoPart Industriesensorik GmbH
        #   Type: Object Detected
        $ 1993 "Object Detected" "noBreak"
        if (visor_partsFound(easyPickVisorId) > 0):
          $ 1994 "Open Gripper" "noBreak"
          # begin: URCap Program Node
          #   Source: Robotiq_Grippers, 1.8.4.4844, Robotiq Inc.
          #   Type: Gripper
          $ 1995 "Gripper Open (1)" "noBreak"
          if not(gripper_connected[0]):
            popup("Gripper 1 must be connected to run this program.", "No connection", False, True, True)
          end
          if not(rq_is_gripper_activated("1")):
            popup("Gripper 1 is not activated. Go to Installation tab > Gripper to activate it and run the program again.", "Not activated", False, True, True)
          end
          rq_set_pos_spd_for(0, 102, 77, "1")
          rq_wait_pos_spe_for_request(0, 102, 77, "1")
          rq_go_to("1")
          rq_wait("1")
          # end: URCap Program Node
          $ 1996 "MoveJ" "noBreak"
          $ 1997 "Waypoint_13" "noBreak"
          movej(get_inverse_kin(Waypoint_13_p, qnear=Waypoint_13_q), a=1.3962634015954636, v=1.0471975511965976)
          # begin: URCap Program Node
          #   Source: SensoPart VISOR Robotic, 2.0.0, SensoPart Industriesensorik GmbH
          #   Type: Approach Pose
          $ 1998 "Approach Pose" "noBreak"
          movej(pose_trans(easyPickPose,p[0.0000,0.0000,0.0500,0.0000,0.0000,0.0000]),a=1.3963,v=1.0472,t=0.000000,r=0.000000)
          # end: URCap Program Node
          # begin: URCap Program Node
          #   Source: SensoPart VISOR Robotic, 2.0.0, SensoPart Industriesensorik GmbH
          #   Type: Target Pose
          $ 1999 "Target Pose" "noBreak"
          movel(pose_trans(easyPickPose,p[0.0000,0.0000,-0.0000,0.0000,0.0000,0.0000]),a=0.5000,v=0.2500,t=0.000000,r=0.000000)
          # end: URCap Program Node
          $ 2000 "Close Gripper" "noBreak"
          # begin: URCap Program Node
          #   Source: Robotiq_Grippers, 1.8.4.4844, Robotiq Inc.
          #   Type: Gripper
          $ 2001 "Gripper Close (1)" "noBreak"
          if not(gripper_connected[0]):
            popup("Gripper 1 must be connected to run this program.", "No connection", False, True, True)
          end
          if not(rq_is_gripper_activated("1")):
            popup("Gripper 1 is not activated. Go to Installation tab > Gripper to activate it and run the program again.", "Not activated", False, True, True)
          end
          rq_set_pos_spd_for(255, 102, 77, "1")
          rq_wait_pos_spe_for_request(255, 102, 77, "1")
          rq_go_to("1")
          rq_wait("1")
          # end: URCap Program Node
          # begin: URCap Program Node
          #   Source: SensoPart VISOR Robotic, 2.0.0, SensoPart Industriesensorik GmbH
          #   Type: Exit Pose
          $ 2002 "Exit Pose" "noBreak"
          movel(pose_trans(easyPickPose,p[0.0000,0.0000,0.0500,0.0000,0.0000,0.0000]),a=0.5000,v=0.2500,t=0.000000,r=0.000000)
          # end: URCap Program Node
          easyPickObjTaken = True
        end
        # end: URCap Program Node
        # begin: URCap Program Node
        #   Source: SensoPart VISOR Robotic, 2.0.0, SensoPart Industriesensorik GmbH
        #   Type: No Object Detected
        $ 2003 "No Object Detected" "noBreak"
        if (visor_partsFound(easyPickVisorId) < 1):
          $ 2004 "Popup: No Container detected" "noBreak"
          popup("No Container detected", "Message", False, False, blocking=True)
          else:
        end
        # end: URCap Program Node
      end
      easyPickCount = easyPickCount + 1
      visor_easyPickUpdate(easyPickVisorId, "counter", easyPickCount)
      visor_easyPickSetIdent("9ca581", easyPickVisorId)
      # end: URCap Program Node
    end
    visorFuncEasyPick_084428()
    # end: URCap Program Node
    $ 2005 "MoveJ"
    $ 2007 "Waypoint_70" "breakAfter"
    movej(get_inverse_kin(Waypoint_70_p, qnear=Waypoint_70_q), a=0.6981317007977318, v=0.5235987755982988)
    $ 2008 "Waypoint_2" "breakAfter"
    movej(get_inverse_kin(Waypoint_2_p, qnear=Waypoint_2_q), a=0.8726646259971648, v=0.5235987755982988, r=0.05)
    $ 2009 "Waypoint_3" "breakAfter"
    movej(get_inverse_kin(Waypoint_3_p, qnear=Waypoint_3_q), a=0.6981317007977318, v=0.5235987755982988, r=0.05)
    $ 2010 "MoveL"
    $ 2011 "Waypoint_15" "breakAfter"
    movel(Waypoint_15_p, a=0.5, v=0.1, r=0.05)
    $ 2012 "Waypoint_14" "breakAfter"
    movel(Waypoint_14_p, a=0.3, v=0.1)
    $ 2013 "Waypoint_4" "breakAfter"
    movel(Waypoint_4_p, a=0.3, v=0.05)
    # begin: URCap Program Node
    #   Source: Robotiq_Grippers, 1.8.4.4844, Robotiq Inc.
    #   Type: Gripper
    $ 2014 "Gripper Open (1)"
    if not(gripper_connected[0]):
      popup("Gripper 1 must be connected to run this program.", "No connection", False, True, True)
    end
    if not(rq_is_gripper_activated("1")):
      popup("Gripper 1 is not activated. Go to Installation tab > Gripper to activate it and run the program again.", "Not activated", False, True, True)
    end
    rq_set_pos_spd_for(0, 102, 77, "1")
    rq_wait_pos_spe_for_request(0, 102, 77, "1")
    rq_go_to("1")
    rq_wait("1")
    # end: URCap Program Node
    $ 2015 "MoveL"
    $ 2016 "Waypoint_25" "breakAfter"
    movel(Waypoint_25_p, a=0.3, v=0.1)
    $ 2017 "Waypoint_15" "breakAfter"
    movel(Waypoint_15_p, a=0.5, v=0.1, r=0.05)
    $ 2018 "Home (Safe)"
    movej([-1.2302089344500047, -1.2969853503591224, -1.875639182904262, -1.539621866126728, 1.5731943360401213, -2.80099559440227], a=1.3962634015954636, v=1.0471975511965976)
  elif (36 == switch_1):
    $ 2048 "Case 36"
    $ 2052 "Decap"
    $ 2090 "MoveJ"
    $ 2091 "Waypoint_39" "breakAfter"
    movej(get_inverse_kin(Waypoint_39_p, qnear=Waypoint_39_q), a=1.3962634015954636, v=1.0471975511965976)
    $ 2092 "MoveL"
    $ 2093 "Waypoint_41" "breakAfter"
    movel(Waypoint_41_p, a=0.5, v=0.1)
    $ 2094 "Waypoint_40" "breakAfter"
    movel(Waypoint_40_p, a=0.3, v=0.05)
    # begin: URCap Program Node
    #   Source: Robotiq_Grippers, 1.8.4.4844, Robotiq Inc.
    #   Type: Gripper
    $ 2095 "Gripper Close (1)"
    if not(gripper_connected[0]):
      popup("Gripper 1 must be connected to run this program.", "No connection", False, True, True)
    end
    if not(rq_is_gripper_activated("1")):
      popup("Gripper 1 is not activated. Go to Installation tab > Gripper to activate it and run the program again.", "Not activated", False, True, True)
    end
    rq_set_pos_spd_for(255, 77, 51, "1")
    rq_wait_pos_spe_for_request(255, 77, 51, "1")
    rq_go_to("1")
    rq_wait("1")
    # end: URCap Program Node
    $ 2096 "Loop 2 times"
    Loop_2 = 0
    while (Loop_2 < 2):
      $ 2097 "MoveL"
      $ 2098 "Waypoint_42" "breakAfter"
      movel(Waypoint_42_p, a=1.2, v=0.5)
      $ 2099 "Waypoint_43" "breakAfter"
      movel(Waypoint_43_p, a=1.2, v=0.25)
      # begin: URCap Program Node
      #   Source: Robotiq_Grippers, 1.8.4.4844, Robotiq Inc.
      #   Type: Gripper
      $ 2100 "Gripper Move40mm (1)"
      if not(gripper_connected[0]):
        popup("Gripper 1 must be connected to run this program.", "No connection", False, True, True)
      end
      if not(rq_is_gripper_activated("1")):
        popup("Gripper 1 is not activated. Go to Installation tab > Gripper to activate it and run the program again.", "Not activated", False, True, True)
      end
      rq_set_pos_spd_for(63, 77, 51, "1")
      rq_wait_pos_spe_for_request(63, 77, 51, "1")
      rq_go_to("1")
      rq_wait("1")
      # end: URCap Program Node
      $ 2101 "MoveL"
      $ 2102 "Waypoint_44" "breakAfter"
      movel(Waypoint_44_p, a=1.2, v=0.5)
      $ 2103 "Waypoint_45" "breakAfter"
      movel(Waypoint_45_p, a=1.2, v=0.25)
      # begin: URCap Program Node
      #   Source: Robotiq_Grippers, 1.8.4.4844, Robotiq Inc.
      #   Type: Gripper
      $ 2104 "Gripper Move11mm (1)"
      if not(gripper_connected[0]):
        popup("Gripper 1 must be connected to run this program.", "No connection", False, True, True)
      end
      if not(rq_is_gripper_activated("1")):
        popup("Gripper 1 is not activated. Go to Installation tab > Gripper to activate it and run the program again.", "Not activated", False, True, True)
      end
      rq_set_pos_spd_for(200, 77, 51, "1")
      rq_wait_pos_spe_for_request(200, 77, 51, "1")
      rq_go_to("1")
      rq_wait("1")
      # end: URCap Program Node
      Loop_2 = Loop_2 + 1
    end
    $ 2105 "MoveL"
    $ 2106 "Waypoint_46" "breakAfter"
    movel(Waypoint_46_p, a=0.3, v=0.05)
    $ 2107 "Waypoint_47" "breakAfter"
    movel(Waypoint_47_p, a=0.5, v=0.1)
    $ 2108 "Waypoint_48" "breakAfter"
    movel(Waypoint_48_p, a=1.2, v=0.25)
    $ 2109 "Waypoint_49" "breakAfter"
    movel(Waypoint_49_p, a=1.2, v=0.25)
    # begin: URCap Program Node
    #   Source: Robotiq_Grippers, 1.8.4.4844, Robotiq Inc.
    #   Type: Gripper
    $ 2110 "Gripper Move35mm (1)"
    if not(gripper_connected[0]):
      popup("Gripper 1 must be connected to run this program.", "No connection", False, True, True)
    end
    if not(rq_is_gripper_activated("1")):
      popup("Gripper 1 is not activated. Go to Installation tab > Gripper to activate it and run the program again.", "Not activated", False, True, True)
    end
    rq_set_pos_spd_for(87, 77, 51, "1")
    rq_wait_pos_spe_for_request(87, 77, 51, "1")
    rq_go_to("1")
    rq_wait("1")
    # end: URCap Program Node
    $ 2111 "MoveL"
    $ 2112 "Waypoint_50" "breakAfter"
    movel(Waypoint_50_p, a=1.2, v=0.25)
    $ 2113 "Home (Safe)"
    movej([-1.2302089344500047, -1.2969853503591224, -1.875639182904262, -1.539621866126728, 1.5731943360401213, -2.80099559440227], a=1.3962634015954636, v=1.0471975511965976)
  elif (37 == switch_1):
    $ 2114 "Case 37"
    $ 2115 "Powder dispensing"
    $ 2116 "zero_scale()"
    zero_scale()
    # begin: URCap Program Node
    #   Source: SensoPart VISOR Robotic, 2.0.0, SensoPart Industriesensorik GmbH
    #   Type: VISOR Robotic App
    $ 2117 "VISOR Easy Pick"
    def visorFuncEasyPick_a4e600():
      # begin: URCap Program Node
      #   Source: SensoPart VISOR Robotic, 2.0.0, SensoPart Industriesensorik GmbH
      #   Type: Easy Pick Setup
      $ 2118 "# 1 Setup" "noBreak"
      local easyPickVisorId = 1
      local easyPickArmMounted = True
      local easyPickSetJob = True
      local easyPickJobName = "Weigh_scale"
      local easyPickAtImgAcq = False
      local easyPickImgAcqPose = cont_img_pose
      # end: URCap Program Node
      # begin: URCap Program Node
      #   Source: SensoPart VISOR Robotic, 2.0.0, SensoPart Industriesensorik GmbH
      #   Type: Process
      $ 2119 "Process" "noBreak"
      local easyPickObjTaken = False
      local easyPickTrigger = False
      local easyPickPoseIdx = 0
      local easyPickPose = p[0,0,0,0,0,0]
      def easyPickFuncTrigger(visorId, setJob, jobName, arm):
      if (setJob):
        visor_changeJob(visorId, jobName, 6000)
      end
      if (arm):
        visor_trigger(visorId, 6000, "arm")
      else:
        visor_trigger(visorId, 6000)
      end
      global easyPickParts_4=visor_partsFound(visorId)
      visor_easyPickUpdate(visorId, "parts", visor_partsFound(visorId))
      return visor_getPose3d(visorId, 0)
    end
    while (not easyPickObjTaken):
      easyPickTrigger = (easyPickCount_4 >= visor_partsFound(easyPickVisorId)) or (easyPickCount_4 > 9) or (not visor_easyPickCheckIdent("b1dffd", easyPickVisorId))
      if (easyPickTrigger):
        easyPickCount_4 = 0
      end
      easyPickPoseIdx = easyPickCount_4
      easyPickPose = visor_getPose3d(easyPickVisorId, easyPickPoseIdx)
      visor_easyPickUpdate(easyPickVisorId, "counter", easyPickPoseIdx)
      # begin: URCap Program Node
      #   Source: SensoPart VISOR Robotic, 2.0.0, SensoPart Industriesensorik GmbH
      #   Type: Image Acquisition Pose
      $ 2120 "Image Acquisition Pose" "noBreak"
      if (easyPickTrigger):
        if (not easyPickAtImgAcq):
          movej(pose_trans(easyPickImgAcqPose,p[0.0000,0.0000,-0.0000,0.0000,0.0000,0.0000]),a=1.3963,v=1.0472,t=0.000000,r=0.000000)
          easyPickAtImgAcq = True
        end
        easyPickPose = easyPickFuncTrigger(easyPickVisorId, easyPickSetJob, easyPickJobName, easyPickArmMounted)
      end
      # end: URCap Program Node
      # begin: URCap Program Node
      #   Source: SensoPart VISOR Robotic, 2.0.0, SensoPart Industriesensorik GmbH
      #   Type: Object Detected
      $ 2121 "Object Detected" "noBreak"
      if (visor_partsFound(easyPickVisorId) > 0):
        $ 2122 "Open Gripper" "noBreak"
        $ 2123 "MoveL" "noBreak"
        $ 2124 "Weight_value≔get_weight()" "noBreak"
        global Weight_value=get_weight()
        # begin: URCap Program Node
        #   Source: Robotiq_Grippers, 1.8.4.4844, Robotiq Inc.
        #   Type: Gripper
        $ 2125 "Gripper Open (1)" "noBreak"
        if not(gripper_connected[0]):
          popup("Gripper 1 must be connected to run this program.", "No connection", False, True, True)
        end
        if not(rq_is_gripper_activated("1")):
          popup("Gripper 1 is not activated. Go to Installation tab > Gripper to activate it and run the program again.", "Not activated", False, True, True)
        end
        rq_set_pos_spd_for(0, 77, 77, "1")
        rq_wait_pos_spe_for_request(0, 77, 77, "1")
        rq_go_to("1")
        rq_wait("1")
        # end: URCap Program Node
        $ 2126 "Waypoint_53" "noBreak"
        movel(Waypoint_53_p, a=0.6, v=0.15, r=0.05)
        $ 2127 "Spatula_above" "noBreak"
        movel(Spatula_above_p, a=0.6, v=0.15)
        $ 2128 "Spatula_pick" "noBreak"
        movel(Spatula_pick_p, a=0.6, v=0.15)
        # begin: URCap Program Node
        #   Source: Robotiq_Grippers, 1.8.4.4844, Robotiq Inc.
        #   Type: Gripper
        $ 2129 "Gripper Close (1)" "noBreak"
        if not(gripper_connected[0]):
          popup("Gripper 1 must be connected to run this program.", "No connection", False, True, True)
        end
        if not(rq_is_gripper_activated("1")):
          popup("Gripper 1 is not activated. Go to Installation tab > Gripper to activate it and run the program again.", "Not activated", False, True, True)
        end
        rq_set_pos_spd_for(255, 77, 77, "1")
        rq_wait_pos_spe_for_request(255, 77, 77, "1")
        rq_go_to("1")
        rq_wait("1")
        # end: URCap Program Node
        $ 2130 "Spatula_above" "noBreak"
        movel(Spatula_above_p, a=0.6, v=0.15)
        $ 2131 "Popup: Connect the vibration motor" "noBreak"
        popup("Connect the vibration motor", "Message", False, False, blocking=True)
        $ 2132 "tare_scale()" "noBreak"
        tare_scale()
        $ 2133 "container_start" "noBreak"
        movel(container_start_p, a=0.3, v=0.1)
        $ 2134 "container_wp_1" "noBreak"
        movel(container_wp_1_p, a=0.3, v=0.05)
        $ 2135 "Loop 1 times" "noBreak"
        Loop_9 = 0
        while (Loop_9 < 1):
          $ 2136 "Waypoint_55" "noBreak"
          global move_thread_flag_2136=0
          thread move_thread_2136():
            enter_critical
            move_thread_flag_2136 = 1
            movel(Waypoint_55_p, a=0.5, v=0.07)
            move_thread_flag_2136 = 2
            exit_critical
          end
          move_thread_flag_2136 = 0
          move_thread_han_2136 = run move_thread_2136()
          while (True):
            sleep(1.0E-10)
            if (move_thread_flag_2136 > 1):
              join move_thread_han_2136
              break
            end
            sync()
          end
          $ 2138 "Waypoint_56" "noBreak"
          movel(Waypoint_56_p, a=0.3, v=0.05)
          $ 2139 "Waypoint_74" "noBreak"
          movel(Waypoint_74_p, a=0.6, v=0.15)
          $ 2140 "Set AO[0]=3.0" "noBreak"
          set_standard_analog_out(0, 0.3)
          $ 2141 "Wait: 2.0" "noBreak"
          sleep(2.0)
          $ 2142 "Set AO[0]=0.0" "noBreak"
          set_standard_analog_out(0, 0.0)
          Loop_9 = Loop_9 + 1
        end
        $ 2146 "ftr_scoop2" "noBreak"
        movel(ftr_scoop2_p, a=0.3, v=0.05)
        $ 2147 "aftr_scoo3" "noBreak"
        movel(aftr_scoo3_p, a=0.3, v=0.05)
        $ 2148 "MoveJ" "noBreak"
        $ 2149 "Waypoint_60" "noBreak"
        movej(get_inverse_kin(Waypoint_60_p, qnear=Waypoint_60_q), a=0.5235987755982988, v=0.3490658503988659, r=0.05)
        $ 2150 "Waypoint_61" "noBreak"
        movej(get_inverse_kin(Waypoint_61_p, qnear=Waypoint_61_q), a=0.5235987755982988, v=0.3490658503988659, r=0.05)
        # begin: URCap Program Node
        #   Source: SensoPart VISOR Robotic, 2.0.0, SensoPart Industriesensorik GmbH
        #   Type: Approach Pose
        $ 2151 "Approach Pose" "noBreak"
        movej(pose_trans(easyPickPose,p[0.0000,0.0000,0.0500,0.0000,0.0000,0.0000]),a=0.4363,v=0.3491,t=0.000000,r=0.000000)
        # end: URCap Program Node
        # begin: URCap Program Node
        #   Source: SensoPart VISOR Robotic, 2.0.0, SensoPart Industriesensorik GmbH
        #   Type: Target Pose
        $ 2152 "Target Pose" "noBreak"
        movel(pose_trans(easyPickPose,p[0.0000,0.0000,-0.0000,0.0000,0.0000,0.0000]),a=0.1000,v=0.0500,t=0.000000,r=0.000000)
        # end: URCap Program Node
        $ 2153 "Close Gripper" "noBreak"
        $ 2154 "dispense_pos≔get_actual_tcp_pose()" "noBreak"
        global dispense_pos= get_actual_tcp_pose ()
        $ 2155 "MoveL" "noBreak"
        $ 2156 "Start_thread≔ True " "noBreak"
        global Start_thread=  True
        $ 2157 "vib_mot_thread≔ True " "noBreak"
        global vib_mot_thread=  True
        $ 2158 "tilt_angle≔current_pose[4]" "noBreak"
        global tilt_angle=current_pose[4]
        $ 2159 "Wait: 0.5" "noBreak"
        sleep(0.5)
        $ 2160 "Loop Weight_value≤Target_weight and tilt_angle≤-0.40" "noBreak"
        thread Thread_while_2160():
          while (True):
            $ 2161 "current_error≔Target_weight-Weight_value" "noBreak"
            global current_error=Target_weight-Weight_value
            $ 2162 "Integral_error≔Integral_error+current_error*dt" "noBreak"
            global Integral_error=Integral_error+current_error*dt
            $ 2163 "derivative≔(current_error-previous_error)/dt" "noBreak"
            global derivative=(current_error-previous_error)/dt
            $ 2164 "tilt_increment≔(kp*current_error)+(ki*Integral_error)+(kd*derivative)" "noBreak"
            global tilt_increment=(kp*current_error)+(ki*Integral_error)+(kd*derivative)
            $ 2165 "current_pose≔get_actual_tcp_pose()" "noBreak"
            global current_pose= get_actual_tcp_pose ()
            $ 2166 "tilt_angle≔current_pose[4]" "noBreak"
            global tilt_angle=current_pose[4]
            $ 2167 "tilt_pose≔pose_trans(current_pose, p[(tilt_increment/7), 0, 0, 0, tilt_increment, 0])" "noBreak"
            global tilt_pose=pose_trans(current_pose, p[(tilt_increment/7), 0, 0, 0, tilt_increment, 0])
            $ 2168 "movel(tilt_pose, a=0.025, v=0.015, r=0.00001)" "noBreak"
            movel(tilt_pose, a=0.025, v=0.015, r=0.00001)
            $ 2169 "previous_error≔current_error" "noBreak"
            global previous_error=current_error
          end
        end
        if (Weight_value <= Target_weight  and  tilt_angle <= -0.40):
          global thread_handler_2160=run Thread_while_2160()
          while (Weight_value <= Target_weight  and  tilt_angle <= -0.40):
            sync()
          end
          kill thread_handler_2160
        end
        $ 2170 "Start_thread≔ False " "noBreak"
        global Start_thread=  False
